  def clear_socket_buffer(gripper_socket="1", read_timeout = 0.1):
      rq_comm_clear_socket_buffer_enabled[rq_socket_to_index(gripper_socket)] = True
  end

  def rq_gripper_id_to_ascii(gripper_id):
      if(gripper_id == "1"):
          return 57
      elif(gripper_id == "2"):
          return 50
      elif(gripper_id == "3"):
          return 51
      elif(gripper_id == "4"):
          return 52
      end
  end

      def scale(value, rawRange, scaledRange):
          def computeSlope(inputRange, outputRange):
              outputRangeDelta = outputRange[1] - outputRange[0]
              inputRangeDelta = inputRange[1] - inputRange[0]

              if (inputRangeDelta == 0):
                  return 0
              else:
                  return outputRangeDelta / inputRangeDelta
              end
          end

          def computeIntercept(slope, inputRange, outputRange):
              return outputRange[0] - (slope * inputRange[0])
          end

          def clipScaledValue(outputScaledValue, outputRange):
              if (outputRange[0] < outputRange[1]):
                  return clipWhenLowerLimitIsLessThanHigher(outputScaledValue, outputRange)
              else:
                  return clipWhenLowerLimitIsGreaterThanHigherLimit(outputScaledValue, outputRange)
              end
          end

          def clipWhenLowerLimitIsGreaterThanHigherLimit(outputScaledValue, outputRange):
              if (outputScaledValue < outputRange[1]):
                  return outputRange[1]
              elif (outputScaledValue > outputRange[0]):
                  return outputRange[0]
              else:
                  return outputScaledValue
              end
          end

          def clipWhenLowerLimitIsLessThanHigher(outputScaledValue, outputRange):
              if (outputScaledValue < outputRange[0]):
                  return outputRange[0]
              elif (outputScaledValue > outputRange[1]):
                  return outputRange[1]
              else:
                  return outputScaledValue
              end
          end

          slope = computeSlope(rawRange, scaledRange)
          intercept = computeIntercept(slope, rawRange, scaledRange)
          scaledValue = slope * value + intercept
          return clipScaledValue(scaledValue, scaledRange)
      end

      def limit(value, range):
          return scale(value, range, range)
      end


  rq_init_comm_if_connected(9, "1")
  rq_init_comm_if_connected(2, "2")
  rq_init_comm_if_connected(3, "3")
  rq_init_comm_if_connected(4, "4")
  rq_print_connected_grippers()
  rq_gripper_communication_thread = run rq_gripper_communication()
  set_closed_norm(97.6470588235294, "1")
  set_open_norm(1.1764705882352942, "1")
  set_closed_mm(0.0, "1")
  set_open_mm(53.0, "1")
  set_closed_norm(100.0, "2")
  set_open_norm(0.0, "2")
  set_closed_mm(0.0, "2")
  set_open_mm(50.0, "2")
  set_closed_norm(100.0, "3")
  set_open_norm(0.0, "3")
  set_closed_mm(0.0, "3")
  set_open_mm(50.0, "3")
  set_closed_norm(100.0, "4")
  set_open_norm(0.0, "4")
  set_closed_mm(0.0, "4")
  set_open_mm(50.0, "4")
  rq_current_limit_enabled = False
  while(not rq_gripper_communication_thread_started):
      sleep(0.008)
  end
  # end: URCap Installation Node
  global AMR_Position=struct(position_identifier=0, x1=0, x2=0, y1=0, y2=0, theta1=0, theta2=0)
  global CAM_Pose=p[0,0,0,0,0,0]
  global CAM_Relation=""
  global CMD_Abort=  False
  global CMD_Clear=  False
  global CMD_Reset=  False
  global CMD_Start=  False
  global CMD_Suspend=  False
  global CMD_Unhold=  False
  global CMD_Unsuspend=  False
  global CNT_Rack_Output=0
  global FNC_Freedrive=  False
  global PRC_TubCounter=0
  global STP=0
  global easyPickCount_4=0
  global easyPickCount_7=0
  global easyPickNoObj_4=0
  global easyPickNoObj_7=0
  global easyPickParts_4=0
  global easyPickParts_7=0
  global TMR_Barcode=0
  global Container_mid_1_p=p[-.379239199143, -.127191311915, .299999999998, .000000000046, -.000000000021, -1.247199999994]
  global Container_mid_1_q=[-2.477408934449926, -1.2969853503591224, -1.875639182904262, -1.539621866126728, 1.5731943360401213, -2.8009955944022717]
  global trigger_otw_p=p[-.364831738276, -.163967193938, .343299997821, .000000000046, -.000000000020, -1.148401333327]
  global trigger_otw_q=[-2.378283213085033, -1.2994862387706814, -1.7634300687554951, -1.6493302004167063, 1.573123683454141, -2.8011223671816943]
  global Waypoint_54_p=p[.008800512419, -.547926542621, .402696567415, -.589884378425, -.007228654778, -.061268144704]
  global Waypoint_54_q=[-1.2044575850116175, -1.3416667741588135, -1.8272563219070435, -0.9884541195682068, 1.3621035814285278, -2.7712565104113978]
  global Waypoint_77_p=p[-.178371829612, -.433927395311, .368082383916, -.086593488055, .704679941724, -.007869906074]
  global Waypoint_77_q=[-1.265390698109762, -1.3355963987163086, -1.7944865226745605, -1.7402602634825648, 0.8780410885810852, -2.7713127771960657]
  global Waypoint_83_p=p[.008800512419, -.547926542621, .402696567415, -.589884378425, -.007228654778, -.061268144704]
  global Waypoint_83_q=[-1.2044575850116175, -1.3416667741588135, -1.8272563219070435, -0.9884541195682068, 1.3621035814285278, -2.7712565104113978]
  global Waypoint_84_p=p[-.178371829612, -.433927395311, .368082383916, -.086593488055, .704679941724, -.007869906074]
  global Waypoint_84_q=[-1.265390698109762, -1.3355963987163086, -1.7944865226745605, -1.7402602634825648, 0.8780410885810852, -2.7713127771960657]
  global Vial_above_1_p=p[.017105793010, -.652093028359, .184920586844, .000000000272, .000000000270, 1.564063451276]
  global Vial_above_1_q=[-1.3375440709712851, -1.9618096977868804, -1.4665759083780685, -1.2837941559171444, 1.5732503672317195, -4.47276330421513]
  global Vial_pick_poi_1_p=p[.017105792852, -.648922724010, .093307568731, .000000000271, .000000000270, 1.564063451276]
  global Vial_pick_poi_1_q=[-1.3366329456391917, -2.0375277831965413, -1.6071432798879028, -1.0675084332049813, 1.57309887265915, -4.471135348858068]
  global Waypoint_86_p=p[.019227646885, -.648669633640, .184920586950, .000000000000, .000000000000, .024063451426]
  global Waypoint_86_q=[-1.3331129109407733, -1.9540750545686123, -1.4775914902901128, -1.280581784992414, 1.5733500744865856, -2.928303704452631]
  global Waypoint_87_p=p[-.032361834699, -.348336136197, .391475576335, -.000008499254, .000014589902, -.004651426820]
  global Waypoint_87_q=[-1.2709335019096129, -1.1914598663441005, -1.708995335060501, -1.8117888533498316, 1.5729683532263925, -2.8379347397710237]
  global Vial_3FG_plac_1_p=p[-.031858676359, -.349402499566, .145301120695, .000000000000, .000000000000, .000000000000]
  global Vial_3FG_plac_1_q=[-1.2723975525801707, -1.252376585823825, -2.3128114007049496, -1.1470592278900167, 1.5730548099411423, -2.8414815174610535]
  global Waypoint_88_p=p[-.032361834699, -.348336136197, .391475576335, -.000008499254, .000014589902, -.004651426820]
  global Waypoint_88_q=[-1.2709335019096129, -1.1914598663441005, -1.708995335060501, -1.8117888533498316, 1.5729683532263925, -2.8379347397710237]
  global cap_dump_1_p=p[-.139168676487, -.420163541420, .146096395183, .000000000000, .000000000000, .000000000000]
  global cap_dump_1_q=[-1.584588644510994, -1.5093464179777323, -2.1118449369620347, -1.091059703602438, 1.5728943834877336, -3.154014906686923]
  global Waypoint_89_p=p[-.032361834699, -.348336136197, .391475576335, -.000008499254, .000014589902, -.004651426820]
  global Waypoint_89_q=[-1.2709335019096129, -1.1914598663441005, -1.708995335060501, -1.8117888533498316, 1.5729683532263925, -2.8379347397710237]
  global Vial_3FG_plac_2_p=p[-.031858676359, -.349402499566, .145301120695, .000000000000, .000000000000, .000000000000]
  global Vial_3FG_plac_2_q=[-1.2723975525801707, -1.252376585823825, -2.3128114007049496, -1.1470592278900167, 1.5730548099411423, -2.8414815174610535]
  global Waypoint_90_p=p[-.032361834699, -.348336136197, .391475576335, -.000008499254, .000014589902, -.004651426820]
  global Waypoint_90_q=[-1.2709335019096129, -1.1914598663441005, -1.708995335060501, -1.8117888533498316, 1.5729683532263925, -2.8379347397710237]
  global cap_dump_2_p=p[-.139168676487, -.420163541420, .146096395183, .000000000000, .000000000000, .000000000000]
  global cap_dump_2_q=[-1.584588644510994, -1.5093464179777323, -2.1118449369620347, -1.091059703602438, 1.5728943834877336, -3.154014906686923]
  global Waypoint_91_p=p[-.032361834699, -.348336136197, .391475576335, -.000008499254, .000014589902, -.004651426820]
  global Waypoint_91_q=[-1.2709335019096129, -1.1914598663441005, -1.708995335060501, -1.8117888533498316, 1.5729683532263925, -2.8379347397710237]
  global Vial_liq_abov_1_p=p[-.025303660977, -.338758622354, .426628485936, -1.315858642253, .800043520260, -.928295855026]
  global Vial_liq_abov_1_q=[-0.3789628187762659, -1.5149522957256814, -2.263045310974121, 0.7870649534412841, -0.750984017048971, -3.2237566153155726]
  global Vial_liq_pick_3_p=p[-.002660428945, -.335984893034, .159389832934, -1.150456778400, .673175527684, -1.010612657503]
  global Vial_liq_pick_3_q=[-0.3660772482501429, -1.4503649038127442, -2.4056053161621094, -1.994692941705221, 0.8039668202400208, -0.2508929411517542]
  global Vial_liq_pick_4_p=p[-.041402486291, -.356791603314, .125395323246, -1.143483969075, .651070210027, -.878721885453]
  global Vial_liq_pick_4_q=[-0.4426233705502476, -1.437252121513727, -2.551930962114307, -1.776528229806984, 0.6562026234073748, -0.43018811960029524]
  global Vial_liq_abov_2_p=p[-.025303660977, -.338758622354, .426628485936, -1.315858642253, .800043520260, -.928295855026]
  global Vial_liq_abov_2_q=[-0.3789628187762659, -1.5149522957256814, -2.263045310974121, 0.7870649534412841, -0.750984017048971, -3.2237566153155726]
  global Liquid_midway_1_p=p[.057575295009, -.583081747994, .306414980749, -1.351675548728, .120935756539, -.096908606303]
  global Liquid_midway_1_q=[-0.895174805318014, -1.7035466633238734, -2.380953073501587, 0.631549521083496, 0.7706599235534668, -2.9455552736865442]
  global shake_3_p=p[.057574880217, -.583085370269, .306422893466, -1.360996190983, -.155555042453, -.438136255921]
  global shake_3_q=[-0.8951800505267542, -1.7035466633238734, -2.380937099456787, 0.6315542894550782, 0.7706599235534669, -2.5394540616517496]
  global shake_4_p=p[.057581636113, -.583090570002, .306439684073, -1.308767904323, .368530312677, .214926493520]
  global shake_4_q=[-0.8951714674579065, -1.7035395107665003, -2.380906343460083, 0.6315504747578125, 0.7706480026245118, -3.3161255787892268]
  global drop_above_3_p=p[.268235025993, -.467784390499, .226219872376, -1.027832627524, -.430841408251, 1.004603115937]
  global drop_above_3_q=[-0.935645882283346, -1.6663371525206507, -2.4252893924713135, 0.41966931402172847, 1.8470635414123535, -3.4600217978106897]
  global drop_above_4_p=p[.219042229014, -.470775657081, .133754190740, -.313004595901, -.344395319364, 1.500564994056]
  global drop_above_4_q=[-1.0601594887284795, -1.70046459045642, -2.0799996233759863, -0.7243227230676759, 1.9429634314685202, -4.115129153870795]
  global liq_tran_3_p=p[.213067510942, -.469567035397, .100231043184, .251862243732, .217902579404, 1.592812335393]
  global liq_tran_3_q=[-0.7789645168037476, -1.822364827406652, -1.8643518410805573, -1.252158963840138, 1.3768134449520435, -3.9328333233290254]
  global drop_above_5_p=p[.219042229014, -.470775657081, .133754190740, -.313004595901, -.344395319364, 1.500564994056]
  global drop_above_5_q=[-1.0601594887284795, -1.70046459045642, -2.0799996233759863, -0.7243227230676759, 1.9429634314685202, -4.115129153870795]
  global Waypoint_92_p=p[.187119460405, -.493959476151, .133754190608, -.313004596540, -.344395317757, 1.500564993991]
  global Waypoint_92_q=[-1.1418328121400876, -1.7310553375189475, -2.033634768766424, -0.772026910513711, 1.958578934631971, -4.201588449364511]
  global liq_tran_4_p=p[.195957706507, -.493022614126, .100231042689, .160718757180, .109807038912, 1.525321508623]
  global liq_tran_4_q=[-0.881740380645474, -1.8244526267589851, -1.865100964490387, -1.1608866323693583, 1.4631433601076713, -3.973915130363038]
  global drop_above_6_p=p[.219042229014, -.470775657081, .133754190740, -.313004595901, -.344395319364, 1.500564994056]
  global drop_above_6_q=[-1.0601594887284795, -1.70046459045642, -2.0799996233759863, -0.7243227230676759, 1.9429634314685202, -4.115129153870795]
  global drop_above_7_p=p[.268235025993, -.467784390499, .226219872376, -1.027832627524, -.430841408251, 1.004603115937]
  global drop_above_7_q=[-0.935645882283346, -1.6663371525206507, -2.4252893924713135, 0.41966931402172847, 1.8470635414123535, -3.4600217978106897]
  global Liquid_midway_2_p=p[.057575295009, -.583081747994, .306414980749, -1.351675548728, .120935756539, -.096908606303]
  global Liquid_midway_2_q=[-0.895174805318014, -1.7035466633238734, -2.380953073501587, 0.631549521083496, 0.7706599235534668, -2.9455552736865442]
  global Vial_drop_abo_1_p=p[.000324902251, -.648569523142, .221894115667, -.873462921366, 1.165852672573, -1.482720593185]
  global Vial_drop_abo_1_q=[-1.0576906334721352, -2.393016994184633, -0.9236232851859159, -2.5729213042279273, 0.7903331288549689, -0.33286325848155585]
  global Vial_liq_drop_1_p=p[.001020867953, -.647659915585, .092915870838, -.834762611599, 1.081942994823, -1.540647900176]
  global Vial_liq_drop_1_q=[-1.0631954168193474, -2.4447642951220825, -1.128811017825127, -2.1983115491972294, 0.8130148661460634, -0.38984988696911316]
  global Vial_drop_abo_2_p=p[.000324902251, -.648569523142, .221894115667, -.873462921366, 1.165852672573, -1.482720593185]
  global Vial_drop_abo_2_q=[-1.0576906334721352, -2.393016994184633, -0.9236232851859159, -2.5729213042279273, 0.7903331288549689, -0.33286325848155585]
  global Spatula_otw_p=p[-.038472058237, -.263141484147, .425351216717, -.000441582511, -.000128175490, 3.034387645854]
  global Spatula_otw_q=[-1.1888947506684495, -1.0083288774886814, -1.7052227056065874, -1.9984805067363443, 1.5730180972985317, 0.48793409320312264]
  global pick_spat_L_abv_p=p[.239059466375, -.067212518441, .280720723617, .000017217488, -.000484427718, 3.106837214660]
  global pick_spat_L_abv_q=[0.292765616142962, -0.8565557553273315, -2.140199892763044, -1.715349495646084, 1.573623142106424, 1.8984976776985687]
  global spat_L_pick_p=p[.242468789885, -.067301915011, .193171208067, .000017217488, -.000484427718, 3.106837214657]
  global spat_L_pick_q=[0.2867414378807389, -0.8600077002089179, -2.3629148016312627, -1.4891831672860159, 1.5737695566221115, 1.8933890858591198]
  global spat_L_lift_p=p[.245402002494, -.067432373551, .289049296496, .000017217490, -.000484427724, 3.106837214657]
  global spat_L_lift_q=[0.2834351187564135, -0.8798320076811592, -2.1119436738532986, -1.7203314352121302, 1.573588313403067, 1.8891054681654005]
  global spat_L_side_p=p[.247133573905, -.017633681797, .289062935631, .000017217490, -.000484427724, 3.106837214657]
  global spat_L_side_q=[0.49719173575848863, -0.8582398211168538, -2.1182130454788215, -1.735610316654931, 1.5735817737572706, 2.1028402698705397]
  global spat_L_up_p=p[.247135508752, -.017665230822, .397130746165, .000017217490, -.000484427724, 3.106837214657]
  global spat_L_up_q=[0.49854946074076967, -0.9346239623559676, -1.808280269374471, -1.969158816463132, 1.5731020084036995, 2.1031742024348157]
  global spat_M_up_p=p[.244670000000, -.112000000000, .420343789747, .000026293990, -.000477463070, 3.067686800857]
  global spat_M_up_q=[0.09097498152209688, -1.0114245603211778, -1.718034632879454, -1.9826932847219538, 1.5730130135866505, 1.734554438783734]
  global spat_M_pick_p=p[.244673518506, -.111985070134, .192299022723, .000043885692, -.000001622442, 3.067686841404]
  global spat_M_pick_q=[0.08868170265231701, -0.9271392933223233, -2.343826449241451, -1.441236864368305, 1.5733923850045939, 1.7345552462242537]
  global spat_S_Up_7_p=p[.243228810603, -.161948321982, .423281604617, .000026293955, -.000477463064, 3.067686800854]
  global spat_S_Up_7_q=[-0.11182322368059516, -1.0716267311491734, -1.6854498186860427, -1.955120134033855, 1.5730106579635699, 1.5317349120701778]
  global spat_S_Pick_4_p=p[.245377020686, -.158668022535, .192285730279, .000026293985, -.000477463062, 3.067686800840]
  global spat_S_Pick_4_q=[-0.10087203759495189, -1.011188488703386, -2.311978084495874, -1.3890267520590838, 1.5735990551056096, 1.5450562970948172]
  global spat_S_Up_8_p=p[.252087445596, -.159242094834, .423281604617, .000026293954, -.000477463070, 3.067686800855]
  global spat_S_Up_8_q=[-0.09804692328730358, -1.0862987822056382, -1.6788706463996483, -1.9470242450550348, 1.5730147401359813, 1.5455107082823842]
  global spat_flatM_up_p=p[.229022666361, -.211442909333, .418634047126, .000026293953, -.000477463083, 3.067686800888]
  global spat_flatM_up_q=[-0.30183372580416545, -1.1157042924275036, -1.6775646144685776, -1.9189678841796578, 1.5730340557943228, 1.341766142011193]
  global spat_flatM_pick_p=p[.241028983327, -.208057297586, .192270533170, .000026293950, -.000477463079, 3.067686800885]
  global spat_flatM_pick_q=[-0.2805687960562633, -1.1003763929487214, -2.271431297337675, -1.3404236887924883, 1.5734924238720627, 1.3653813047742556]
  global spat_flatS_up_p=p[.237651953780, -.253943828614, .403961222825, .000026293950, -.000477463092, 3.067686800841]
  global spat_flatS_up_q=[-0.42363550926974103, -1.1939944599502539, -1.6745915127240307, -1.843675057902054, 1.5731001874678698, 1.220082820532415]
  global spat_flatS_pick_p=p[.241325662334, -.251726327528, .192256842740, .000026293947, -.000477463087, 3.067686800841]
  global spat_flatS_pick_q=[-0.4144907797170738, -1.1967447109013012, -2.21926362252748, -1.2962499335425761, 1.5733885098427622, 1.2314402238866728]
  global spat_S_pick_p=p[.238158866340, -.157926795425, .192632100345, .000026293989, -.000477463069, 3.067686800857]
  global spat_S_pick_q=[-0.10084756991493293, -0.9881392730064915, -2.3204232610157494, -1.403630829593915, 1.5736254260650586, 1.5450653591083503]
  global spat_S_up_p=p[.244260523725, -.164466690315, .417087579736, .000026293988, -.000477463072, 3.067686800857]
  global spat_S_up_q=[-0.12101499604198729, -1.0718307017854336, -1.7023391702814736, -1.938028805938881, 1.573044424728474, 1.5226045951991447]
  global Waypoint_7_p=p[-.472820924474, .292439826233, .207418370237, -.137787250486, 2.177332259632, -2.152029714756]
  global Waypoint_7_q=[-2.911134078210732, -1.90240864358569, -1.968768330510411, -2.500365101593811, 0.11427687110891149, 0.0958980389250167]
  global Waypoint_8_p=p[-.357612884176, -.251084817998, .212379799667, -.858181193174, 1.714832512191, -1.687547565568]
  global Waypoint_8_q=[-1.620834863369681, -1.8936194567376496, -1.9821394403832038, -2.4599791457905273, 0.6296693672615152, 0.07625365420707819]
  global Decapp_above_3_p=p[-.013480295948, -.359153355979, .266194408367, -.879653555922, 1.646336924805, -1.709111068605]
  global Decapp_above_3_q=[-0.9632157249872035, -2.0163405763031657, -1.5968194594157152, -2.6579215719847085, 1.251243398585566, 0.047906446502667066]
  global Decapp_place_3_p=p[-.013480295890, -.359153356055, .160907502384, -.879653554902, 1.646336919740, -1.709111066456]
  global Decapp_place_3_q=[-0.9633402410919709, -2.1541179572356635, -1.6937729380888573, -2.4232786481058053, 1.2517342187662468, 0.04818402956922263]
  global Decapp_above_4_p=p[-.013480295948, -.359153355979, .266194408367, -.879653555922, 1.646336924805, -1.709111068605]
  global Decapp_above_4_q=[-0.9632157249872035, -2.0163405763031657, -1.5968194594157152, -2.6579215719847085, 1.251243398585566, 0.047906446502667066]
  global Waypoint_78_p=p[-.051450028091, -.519555688329, .365718563414, -1.287302938145, 1.077637394477, -1.218524965834]
  global Waypoint_78_q=[-0.9214276262416012, -1.8899696965062578, -1.4939326452510562, -2.840015661555725, 0.5585157189668353, 0.033997638875617575]
  global Waypoint_10_p=p[-.330595116596, .282932669854, .220236276291, 1.304675539882, .014233792938, -1.753932442581]
  global Waypoint_10_q=[-3.189526379253601, -1.8418198435143305, -1.7138504750370807, -2.182789974066381, 1.0126080912871243, -2.4455984844694645]
  global Waypoint_9_p=p[-.538777454962, .370695704977, .175030018143, -.317104215445, 2.082346543003, -2.037631421082]
  global Waypoint_9_q=[-3.1158871966457857, -1.998548595120492, -1.941797010061462, -2.2703530575838844, -0.27573365931009164, -0.06926782177267654]
  global Powder_wayp1_p=p[-.472820924474, .292439826233, .207418370237, -.137787250486, 2.177332259632, -2.152029714756]
  global Powder_wayp1_q=[-2.911134078210732, -1.90240864358569, -1.968768330510411, -2.500365101593811, 0.11427687110891149, 0.0958980389250167]
  global Waypoint_2_p=p[-.357612884176, -.251084817998, .212379799667, -.858181193174, 1.714832512191, -1.687547565568]
  global Waypoint_2_q=[-1.620834863369681, -1.8936194567376496, -1.9821394403832038, -2.4599791457905273, 0.6296693672615152, 0.07625365420707819]
  global Postions_otw_p=p[-.010896578244, -.533368729951, .288851175116, -1.233738470894, 1.195331112012, -1.207314088469]
  global Postions_otw_q=[-0.898791023514228, -2.078490033037677, -1.4499891355755317, -2.7624416226992476, 0.6570218891920963, 0.02136606178275929]
  global cont_A_otw_p=p[.070238108556, -.655257851554, .184611566008, -1.090601381517, 1.404822685081, -1.413645380264]
  global cont_A_otw_q=[-0.990969136335913, -2.7123780097559784, -0.5772671651193146, -3.0005537851220403, 0.84719335943793, 0.020652463706785973]
  global cont_B_otw_p=p[.255895686750, -.501120003087, .157855243207, -1.209177187561, 1.209243088037, -1.209202949417]
  global cont_B_otw_q=[-0.5819602570351563, -2.5181180937953833, -1.0264696604583161, -2.7360726814058687, 0.9880932038785559, -0.004134033524621827]
  global cont_B_safe_p=p[.242897168204, -.501733713795, .237745474779, -1.209212324107, 1.209144328638, -1.209309913894]
  global cont_B_safe_q=[-0.5929699566143585, -2.4210115429142114, -0.9949203644592259, -2.8646436479104267, 0.976678899749076, -0.004020526358775811]
  global cont_C_otw_p=p[.319495487998, -.362719410364, .163846736977, -1.233784872294, 1.195277203291, -1.207325031551]
  global cont_C_otw_q=[-0.3611889651645974, -2.404603865546651, -1.2341573845076566, -2.650535279811077, 1.1944844573128257, 0.01638086594640864]
  global Waypoint_1_p=p[-.352029261722, -.424157832422, .472326578019, -.000004407962, .000020663369, -1.529709227737]
  global Waypoint_1_q=[-2.017015745614491, -1.7423968528991196, -1.0053357238485425, -1.9644715035904907, 1.5727249689896, -2.060727852912713]
  global Waypoint_5_p=p[.219993437017, -.447144142811, .462350040687, .000006087494, .000031090075, .000022232405]
  global Waypoint_5_q=[-0.8406239476037944, -1.5982534362206806, -1.1934200873248484, -1.9205794898315975, 1.5727336676986443, -2.4135960466995314]
  global place_2_home_p=p[-.352029261717, -.424157832411, .329197314759, -.000004407962, .000020663369, -1.529709227737]
  global place_2_home_q=[-2.017880982348384, -1.6708952803108668, -1.462293789471877, -1.5790150659586653, 1.5732060241635952, -2.059940179665328]
  global PosA_up_p=p[.028578953747, -.638006009765, .227275735849, -1.090660933958, 1.404791542934, -1.413645191233]
  global PosA_up_q=[-1.0254743496427432, -2.565176838504783, -0.7558042274983681, -2.9696064674274343, 0.8129191411995651, 0.021444818458024387]
  global PosA_pick_p=p[.026918718687, -.640084889741, .097901147521, -1.090660933959, 1.404791542934, -1.413645191233]
  global PosA_pick_q=[-1.028821435558534, -2.6899890636403807, -0.8526126047665157, -2.7478942693937167, 0.8103607002888742, 0.021326778146411485]
  global PosB_up_p=p[.239472634782, -.492481416782, .220767759213, -1.233738470883, 1.195331111998, -1.207314088469]
  global PosB_up_q=[-0.5800230603397054, -2.4076296700885997, -1.0699783327330836, -2.8116344407747427, 0.9750472858169287, 0.017627507888886562]
  global PosB_pick_p=p[.240630296955, -.494558620171, .096392895280, -1.233740573549, 1.195309876041, -1.207293779132]
  global PosB_pick_q=[-0.5816146260408139, -2.553273721769836, -1.1376320925804277, -2.5983292591462153, 0.9740936784345416, 0.017625262979849232]
  global PosC_up_p=p[.241566602786, -.359249123455, .230260583862, -1.233738470888, 1.195331111997, -1.207314088449]
  global PosC_up_q=[-0.39573787962534546, -2.2019009616581497, -1.4115270142506517, -2.675987785326166, 1.160180741930842, 0.01687917643039505]
  global PosC_pick_p=p[.240633854030, -.361553124916, .093979792658, -1.233738470878, 1.195331111997, -1.207314088469]
  global PosC_pick_q=[-0.39992427526118757, -2.386042391328985, -1.4894374567278712, -2.414022930893381, 1.1566786195951169, 0.01712017454263659]
  global Pow_decap_up_p=p[-.017556487132, -.367519866742, .275835445416, -.605635182849, 1.892518157522, -1.890848751165]
  global Pow_decap_up_q=[-1.1272088681128203, -2.1173924123331025, -1.4250048354055203, -2.7485980486387676, 1.4193896902217862, 0.023247957637719453]
  global pow_decap_place_p=p[-.020433194420, -.368310202914, .161281291611, -.605635182838, 1.892518157522, -1.890848751163]
  global pow_decap_place_q=[-1.132360890531647, -2.2521863255983092, -1.5302136899970318, -2.5086176644751683, 1.4149282844269635, 0.02347140074572661]
  global Decap_above_p=p[-.031863883354, -.349974838955, .288042264213, .000000000000, .000000000000, .000000000000]
  global Decap_above_q=[-1.271900116540503, -1.1670201114602632, -1.989291655468758, -1.5559360538518163, 1.573255119759632, -2.842476569674073]
  global Decapp_p=p[-.031864263150, -.349974612700, .230259377740, .000000000000, .000000000000, .000000000000]
  global Decapp_q=[-1.2723555431601419, -1.1810456878410935, -2.1291754890757737, -1.4020263844320349, 1.5732701843074919, -2.842325632263757]
  global Cap_above_p=p[-.224192409203, -.629599568633, .257274081142, .000015605575, -.000015166009, -1.647823825902]
  global Cap_above_q=[-1.710642681834492, -1.9674285251810462, -1.2705185053146897, -1.4742193161331247, 1.573506065067499, -1.6347709465008595]
  global Cap_place_p=p[-.224189049846, -.629597879697, .041885651757, .000015605572, -.000015166011, -1.647823825903]
  global Cap_place_q=[-1.7111696563854295, -2.13979870939016, -1.5941008764912503, -0.978265561728648, 1.5732789016410962, -1.6336328794662904]
  global OP_PowderA2_p=p[.009371277507, -.409434369247, .294169017766, -.823281033205, 1.709410851243, -1.698303593897]
  global OP_PowderA2_q=[-0.9994544761745754, -2.1395254572673217, -1.3437567783153916, -2.8143375616690456, 1.2617899549595724, 0.019614613715634555]
  global Decap_up_p=p[-.018339217391, -.367674469480, .249553854268, -.546164737599, 1.935964719000, -1.930057109666]
  global Decap_up_q=[-1.158124747223252, -2.1569920012936787, -1.4340832185069745, -2.7006032680036753, 1.4556626828962336, 0.02060977878679182]
  global Decap_pick_p=p[-.020429098827, -.367971872627, .161604333799, -.546164737600, 1.935964719000, -1.930057109666]
  global Decap_pick_q=[-1.161653098289774, -2.263509236689538, -1.5087211318402236, -2.519459740767391, 1.452646640403743, 0.02077912034002202]
  global Op_PowA_wP_p=p[-.173727579245, -.372934016396, .295116627479, -.972390492433, 1.540962074418, -1.548745344994]
  global Op_PowA_wP_q=[-1.1740587397768483, -1.865656321049359, -1.7426943793777419, -2.679427276872525, 0.8588908769087338, 0.017944699631825187]
  global Waypoint_12_p=p[-.812560029877, -.415067232840, .258518340146, -1.257569567036, 1.159670338548, -1.145019586130]
  global Waypoint_12_q=[-2.3224548809497123, -2.3211405271930765, -1.1304722687551445, -2.8155296475017018, -0.8321758827962036, -0.007205995478960503]
  global Waypoint_18_p=p[-.813643087636, -.416224939441, .090971414301, -1.257570310932, 1.159676546329, -1.145010619026]
  global Waypoint_18_q=[-2.3224916967547475, -2.513993544062452, -1.2408975037093848, -2.5121717481246186, -0.831286599209303, -0.007326414722441221]
  global Waypoint_19_p=p[-.812560029269, -.415067232191, .079455005744, -1.257569567033, 1.159670338546, -1.145019586137]
  global Waypoint_19_q=[-2.3224951834453367, -2.5274729453886575, -1.2489176533831348, -2.4906644180980346, -0.8312252662037514, -0.007338111970053518]
  global TMR_Barcode_is_counting=False
  thread Timer_Thread():
    while (True):
      if (TMR_Barcode_is_counting):
        TMR_Barcode = TMR_Barcode + get_steptime()
      end
      sync()
    end
  end
  run Timer_Thread()
  def Sub_Vision_V18():
    $ 847 "Sub_Vision_V18" "noBreak"
    $ 848 "PreSettings"
    $ 849 "CAM_LM_Detected≔ False "
    global CAM_LM_Detected=  False
    $ 850 "CAM_Captures≔0"
    global CAM_Captures=0
    $ 851 "CAM_Pose≔p[0,0,0,0,0,0]"
    global CAM_Pose=p[0,0,0,0,0,0]
    $ 852 "CAM_LM_Refinmnt≔ False "
    global CAM_LM_Refinmnt=  False
    $ 853 "CAM_LM_Refined≔ False "
    global CAM_LM_Refined=  False
    $ 854 "CAM_LM_Deviatn≔p[0,0,0,0,0,0]"
    global CAM_LM_Deviatn=p[0,0,0,0,0,0]
    $ 855 "CAM_LM_ID≔0"
    global CAM_LM_ID=0
    $ 856 "CAM_Done≔ False "
    global CAM_Done=  False
    $ 857 "CAM_CNT_Obj≔0"
    global CAM_CNT_Obj=0
    $ 858 "CAM_Result = []"
    CAM_Result = []
    $ 859 "OBJ_Detected≔ False "
    global OBJ_Detected=  False
    $ 860 "FRM_Reference≔p[0,0,0,0,0,0]"
    global FRM_Reference=p[0,0,0,0,0,0]
    $ 861 "'=========='"
    # '=========='
    $ 862 "Switch Action"
    switch_1 = Action
    $ 863 "Case 13"
    if (13 == switch_1):
    elif (15 == switch_1):
      $ 981 "Case 15"
    elif (131 == switch_1):
      $ 1027 "Case 131"
      $ 1028 "Read (SensoPart)"
      $ 1029 "Action_Info≔'search for landmark'"
      global Action_Info="search for landmark"
      $ 1030 "CAM_LM≔CAM_LMs[4]"
      global CAM_LM=CAM_LMs[4]
      $ 1031 "CAM_Relation≔CAM_LM.capture_relation"
      global CAM_Relation=CAM_LM.capture_relation
      $ 1032 "go to capture pose"
      $ 1035 "If ITM_ID≟1 and JIG≟7"
      if (ITM_ID == 1  and  JIG == 7):
        $ 1036 "PSE_T≔uLM_Cap_SSRack"
        global PSE_T=uLM_Cap_SSRack
      else:
        $ 1037 "ElseIf ITM_ID≟5 and JIG≟7"
        if (ITM_ID == 5  and  JIG == 7):
          $ 1038 "PSE_T≔FRM_Cap_SSRack"
          global PSE_T=FRM_Cap_SSRack
        else:
          $ 1041 "ElseIf ITM_ID≟1 and JIG≟15"
          if (ITM_ID == 1 and JIG == 15):
            $ 1042 "MoveJ"
            $ 1043 "Container_mid_1" "breakAfter"
            movej(get_inverse_kin(Container_mid_1_p, qnear=Container_mid_1_q), a=1.3962634015954636, v=1.0471975511965976, r=0.05)
            $ 1045 "PSE_T≔FRM_Container_const"
            global PSE_T=p[-0.5003348223692186,0.35061804815168285,0.41579001388808423,-5.092943187272062E-5,1.0145185065363121E-4,-2.764319258713288]
          else:
            $ 1046 "ElseIf ITM_ID≟1 and JIG≟21"
            if (ITM_ID == 1 and JIG == 21):
              $ 1048 "PSE_T≔FRM_PoTS_const"
              global PSE_T=p[-0.5403054403210852,-0.10910773999775857,0.4828,3.058497512721046E-6,2.3454853329357316E-5,-2.208510541952706]
            else:
              $ 1049 "ElseIf ITM_ID≟1 and JIG≟17"
              if (ITM_ID == 1 and JIG == 17):
                $ 1050 "MoveJ"
                $ 1051 "zero_scale()"
                zero_scale()
                $ 1052 "trigger_otw" "breakAfter"
                movej(get_inverse_kin(trigger_otw_p, qnear=trigger_otw_q), a=1.3962634015954636, v=1.0471975511965976, r=0.05)
                $ 1056 "PSE_T≔FRM_weigh_scale_const"
                global PSE_T=p[-0.3804866881697204,0.025744252835212,0.4723487455232425,-1.0445769542396123E-4,-1.924788411074358E-5,-2.1691978730572363]
              end
            end
          end
        end
      end
      $ 1057 "do_transition(PSE_T, keep_rxry=False)"
      do_transition(PSE_T, keep_rxry=False)
      $ 1058 "Set"
      set_tcp(p[0.0,0.0,0.161,3.1415,0.0,0.0])
      $ 1059 "MoveJ"
      $ 1060 "PSE_T" "breakAfter"
      movej(PSE_T, a=1.3962634015954636, v=1.7453292519943295)
      $ 1061 "CAM_Pose≔get_actual_tcp_pose()"
      global CAM_Pose= get_actual_tcp_pose ()
      $ 1062 "Loop  not CAM_Done and  not ERROR.FLAG and  not CMD_Stop"
      while (  not  CAM_Done  and    not  ERROR.FLAG  and    not  CMD_Stop):
        $ 1063 "adjust capture pose"
        $ 1064 "If CAM_LM_Detected and CAM_LM_Refinmnt"
        if (CAM_LM_Detected  and  CAM_LM_Refinmnt):
          $ 1065 "PSE_T≔p[0,0,0.300,0,0,0]"
          global PSE_T=p[0,0,0.300,0,0,0]
          $ 1066 "CAM_Pose≔PSE_T"
          global CAM_Pose=PSE_T
          $ 1067 "If  not is_reachable(FRM_Reference,[PSE_T])"
          if (  not  is_reachable(FRM_Reference,[PSE_T])):
            $ 1068 "Error"
            $ 1069 "set_error(ERROR_POSE_NOT_REACHABLE)"
            set_error(ERROR_POSE_NOT_REACHABLE)
          end
          $ 1070 "If  not ERROR.FLAG"
          if (  not  ERROR.FLAG):
            $ 1071 "MoveJ"
            $ 1072 "PSE_T" "breakAfter"
            set_tcp(p[0.0,0.0,0.161,0.0,0.0,0.0])
            movej(pose_trans(FRM_Reference, PSE_T), a=0.8726646259971648, v=1.3962634015954636)
            $ 1073 "CAM_LM_Refined≔ True "
            global CAM_LM_Refined=  True
          end
        else:
          $ 1074 "ElseIf  not CAM_LM_Detected and CAM_Captures>0"
          if (  not  CAM_LM_Detected  and  CAM_Captures>0):
            $ 1075 "MoveL"
            $ 1076 "If FRM_Reference≟p[0,0,0,0,0,0]"
            if (FRM_Reference == p[0,0,0,0,0,0]):
              $ 1077 "PSE_T≔get_random_pose(pose_ref=CAM_Pose, mode='cubic', range_max=[0.150,0.150,0.015])"
              global PSE_T=get_random_pose(pose_ref=CAM_Pose, mode="cubic", range_max=[0.150,0.150,0.015])
            else:
              $ 1082 "Else" "noBreak"
              $ 1083 "PSE_T≔get_random_pose(pose_ref=CAM_Pose, mode='rotation', range_max=[10,10,0])"
              global PSE_T=get_random_pose(pose_ref=CAM_Pose, mode="rotation", range_max=[10,10,0])
              $ 1084 "CAM_LM_Refined≔ True "
              global CAM_LM_Refined=  True
            end
            $ 1085 "If get_inverse_kin_has_solution(pose_trans(FRM_Reference, PSE_T))"
            if (get_inverse_kin_has_solution( pose_trans (FRM_Reference, PSE_T))):
              $ 1086 "Comment"
              # Comment
              $ 1087 "PSE_T" "breakAfter"
              set_tcp(p[0.0,0.0,0.161,3.1415,0.0,0.0])
              movel(pose_trans(FRM_Reference, PSE_T), a=0.03, v=0.05)
            else:
              $ 1088 "Else" "noBreak"
              $ 1089 "'If random pose is out of reach, set the initial cam pose'"
              # 'If random pose is out of reach, set the initial cam pose'
              $ 1090 "PSE_T≔CAM_Pose"
              global PSE_T=CAM_Pose
            end
          end
        end
        $ 1091 "Wait: 2.0"
        sleep(2.0)
        $ 1092 "trigger"
        $ 1093 "If ITM_ID≟1 and JIG≟7"
        if (ITM_ID == 1  and  JIG == 7):
          # begin: URCap Program Node
          #   Source: SensoPart VISOR Robotic, 2.0.6, SensoPart Industriesensorik GmbH
          #   Type: VISOR Trigger
          $ 1094 "# 1 VISOR Trigger"
          visor_changeJob(1, "Landmark_INVITE_2", 6000)
          visor_trigger(1, 6000, "arm")
          # end: URCap Program Node
        else:
          $ 1095 "ElseIf ITM_ID≟5 and JIG≟7"
          if (ITM_ID == 5  and  JIG == 7):
            # begin: URCap Program Node
            #   Source: SensoPart VISOR Robotic, 2.0.6, SensoPart Industriesensorik GmbH
            #   Type: VISOR Trigger
            $ 1096 "# 1 VISOR Trigger"
            visor_changeJob(1, "Landmark_INVITE_2", 6000)
            visor_trigger(1, 6000, "arm")
            # end: URCap Program Node
          else:
            $ 1097 "ElseIf ITM_ID≟13 and JIG≟7"
            if (ITM_ID == 13  and  JIG == 7):
              # begin: URCap Program Node
              #   Source: SensoPart VISOR Robotic, 2.0.6, SensoPart Industriesensorik GmbH
              #   Type: VISOR Trigger
              $ 1098 "# 1 VISOR Trigger"
              visor_changeJob(1, "Landmark_INVITE_2", 6000)
              visor_trigger(1, 6000, "arm")
              # end: URCap Program Node
            else:
              $ 1099 "ElseIf ITM_ID≟1 and JIG≟15"
              if (ITM_ID == 1 and JIG == 15):
                # begin: URCap Program Node
                #   Source: SensoPart VISOR Robotic, 2.0.6, SensoPart Industriesensorik GmbH
                #   Type: VISOR Trigger
                $ 1100 "# 1 VISOR Trigger"
                visor_changeJob(1, "Aztec_no_dot_pick", 6000)
                visor_trigger(1, 6000, "arm")
                # end: URCap Program Node
              else:
                $ 1101 "ElseIf ITM_ID≟1 and JIG≟21"
                if (ITM_ID == 1 and JIG == 21):
                  # begin: URCap Program Node
                  #   Source: SensoPart VISOR Robotic, 2.0.6, SensoPart Industriesensorik GmbH
                  #   Type: VISOR Trigger
                  $ 1102 "# 1 VISOR Trigger"
                  visor_changeJob(1, "PoTS", 6000)
                  visor_trigger(1, 6000, "arm")
                  # end: URCap Program Node
                else:
                  $ 1103 "ElseIf ITM_ID≟1 and JIG≟17"
                  if (ITM_ID == 1 and JIG == 17):
                    # begin: URCap Program Node
                    #   Source: SensoPart VISOR Robotic, 2.0.6, SensoPart Industriesensorik GmbH
                    #   Type: VISOR Trigger
                    $ 1104 "# 1 VISOR Trigger"
                    visor_changeJob(1, "Weigh_target", 6000)
                    visor_trigger(1, 6000, "arm")
                    # end: URCap Program Node
                  end
                end
              end
            end
          end
        end
        $ 1108 "TM_3D_Found≔visor_partsFound(1)"
        global TM_3D_Found= visor_partsFound (1)
        $ 1110 "If TM_3D_Found>0"
        if (TM_3D_Found>0):
          $ 1111 "CAM_LM_Detected≔ True "
          global CAM_LM_Detected=  True
          $ 1112 "CAM_Captures≔0"
          global CAM_Captures=0
        else:
          $ 1113 "Else" "noBreak"
          $ 1114 "CAM_LM_Detected≔ False "
          global CAM_LM_Detected=  False
          $ 1115 "CAM_Captures≔CAM_Captures+1"
          global CAM_Captures=CAM_Captures+1
        end
        $ 1120 "result"
        $ 1121 "If CAM_LM_Detected"
        if (CAM_LM_Detected):
          $ 1122 "If (CAM_LM_Refinmnt and CAM_LM_Refined) or  not CAM_LM_Refinmnt"
          if ((CAM_LM_Refinmnt  and  CAM_LM_Refined)  or    not  CAM_LM_Refinmnt):
            $ 1180 "If ITM_ID≟1 and JIG≟7"
            if (ITM_ID == 1  and  JIG == 7):
              $ 1181 "CAM_LM_SSRack≔visor_getPose3d(1, 0)"
              global CAM_LM_SSRack= visor_getPose3d (1, 0)
            else:
              $ 1182 "ElseIf ITM_ID≟5 and JIG≟7"
              if (ITM_ID == 5  and  JIG == 7):
                $ 1183 "CAM_LM_SSRack≔visor_getPose3d(1, 0)"
                global CAM_LM_SSRack= visor_getPose3d (1, 0)
              else:
                $ 1186 "ElseIf ITM_ID≟1 and JIG≟15"
                if (ITM_ID == 1 and JIG == 15):
                  $ 1187 "CAM_LM_cont≔visor_getPose3d(1, 0)"
                  global CAM_LM_cont= visor_getPose3d (1, 0)
                  $ 1188 "Trigger≔get_actual_tcp_pose()"
                  global Trigger= get_actual_tcp_pose ()
                else:
                  $ 1189 "ElseIf ITM_ID≟1 and JIG≟21"
                  if (ITM_ID == 1 and JIG == 21):
                    $ 1190 "CAM_LM_cont≔visor_getPose3d(1, 0)"
                    global CAM_LM_cont= visor_getPose3d (1, 0)
                    $ 1191 "Trigger≔get_actual_tcp_pose()"
                    global Trigger= get_actual_tcp_pose ()
                  else:
                    $ 1192 "ElseIf ITM_ID≟1 and JIG≟17"
                    if (ITM_ID == 1 and JIG == 17):
                      $ 1193 "CAM_LM_cont≔visor_getPose3d(1, 0)"
                      global CAM_LM_cont= visor_getPose3d (1, 0)
                      $ 1194 "Trigger≔get_actual_tcp_pose()"
                      global Trigger= get_actual_tcp_pose ()
                    end
                  end
                end
              end
            end
            $ 1195 "CAM_Done≔ True "
            global CAM_Done=  True
          end
        else:
          $ 1196 "ElseIf  not CAM_LM_Detected and CAM_Captures<CAM_PRM_Retries"
          if (  not  CAM_LM_Detected  and  CAM_Captures<CAM_PRM_Retries):
            $ 1197 "CAM_LM_Refined≔ False "
            global CAM_LM_Refined=  False
          else:
            $ 1198 "ElseIf CAM_Captures≥CAM_PRM_Retries"
            if (CAM_Captures >= CAM_PRM_Retries):
              $ 1199 "CAM_Done≔ True "
              global CAM_Done=  True
              $ 1200 "Error"
              $ 1201 "set_error(ERROR_NO_LANDMARK)"
              set_error(ERROR_NO_LANDMARK)
            end
          end
        end
      end
    elif (151 == switch_1):
      $ 1202 "Case 151"
      $ 1203 "Detect (SensoPart)"
      $ 1204 "go to capture pose"
      $ 1205 "FRM_Reference≔FRM_Cap_SSRack"
      global FRM_Reference=FRM_Cap_SSRack
      $ 1206 "PSE_T≔p[0,0,-0.00,0,0,0]"
      global PSE_T=p[0,0,-0.00,0,0,0]
      $ 1207 "do_transition(pose_trans(FRM_Reference, PSE_T), keep_rxry=False)"
      do_transition( pose_trans (FRM_Reference, PSE_T), keep_rxry=False)
      $ 1208 "JNT_Q≔get_actual_joint_positions()"
      global JNT_Q= get_actual_joint_positions ()
      $ 1209 "JNT_Q≔[JNT_Q[0], JNT_Q[1], JNT_Q[2], JNT_Q[3], JNT_Q[4], 0]"
      global JNT_Q=[JNT_Q[0], JNT_Q[1], JNT_Q[2], JNT_Q[3], JNT_Q[4], 0]
      $ 1210 "Set"
      set_tcp(p[0.0,0.0,0.161,3.1415,0.0,0.0])
      $ 1211 "movej(get_inverse_kin(pose_trans(FRM_Reference, PSE_T), qnear=JNT_Q))"
      movej(get_inverse_kin( pose_trans (FRM_Reference, PSE_T), qnear=JNT_Q))
      $ 1212 "CAM_Pose≔pose_trans(pose_inv(FRM_Reference), get_actual_tcp_pose())"
      global CAM_Pose= pose_trans ( pose_inv (FRM_Reference),  get_actual_tcp_pose ())
      $ 1213 "Loop  not CAM_Done and  not ERROR.FLAG and  not CMD_Stop"
      while (  not  CAM_Done  and    not  ERROR.FLAG  and    not  CMD_Stop):
        $ 1214 "If  not OBJ_Detected and CAM_Captures>0"
        if (  not  OBJ_Detected  and  CAM_Captures>0):
          $ 1215 "MoveL"
          $ 1216 "If FRM_Reference≟p[0,0,0,0,0,0]"
          if (FRM_Reference == p[0,0,0,0,0,0]):
            $ 1218 "PSE_T≔get_random_pose(pose_ref=CAM_Pose, mode='rotation', range_max=[15,15,0])"
            global PSE_T=get_random_pose(pose_ref=CAM_Pose, mode="rotation", range_max=[15,15,0])
          else:
            $ 1219 "Else" "noBreak"
            $ 1220 "PSE_T≔get_random_pose(pose_ref=CAM_Pose, mode='rotation', range_max=[10,10,0])"
            global PSE_T=get_random_pose(pose_ref=CAM_Pose, mode="rotation", range_max=[10,10,0])
          end
          $ 1221 "If get_inverse_kin_has_solution(pose_trans(FRM_Reference, PSE_T))"
          if (get_inverse_kin_has_solution( pose_trans (FRM_Reference, PSE_T))):
            $ 1222 "PSE_T" "breakAfter"
            set_tcp(p[0.0,0.0,0.161,3.1415,0.0,0.0])
            movel(pose_trans(FRM_Reference, PSE_T), a=0.03, v=0.05)
          else:
            $ 1223 "Else" "noBreak"
            $ 1224 "'If random pose is out of reach, set the initial cam pose'"
            # 'If random pose is out of reach, set the initial cam pose'
            $ 1225 "PSE_T≔CAM_Pose"
            global PSE_T=CAM_Pose
            $ 1226 "PSE_T" "breakAfter"
            set_tcp(p[0.0,0.0,0.161,3.1415,0.0,0.0])
            movel(pose_trans(FRM_Reference, PSE_T), a=0.03, v=0.05)
          end
        end
        $ 1227 "Wait: 0.5"
        sleep(0.5)
        $ 1228 "Set"
        set_tcp(p[0.0,0.0,0.161,3.1415,0.0,0.0])
        # begin: URCap Program Node
        #   Source: SensoPart VISOR Robotic, 2.0.6, SensoPart Industriesensorik GmbH
        #   Type: VISOR Trigger
        $ 1229 "# 1 VISOR Trigger"
        visor_changeJob(1, "Object Detection Single", 6000)
        visor_trigger(1, 6000, "arm")
        # end: URCap Program Node
        $ 1230 "If visor_isResponseOk(1)"
        if ( visor_isResponseOk (1)):
          $ 1231 "CAM_CNT_Obj≔visor_partsFound(1)"
          global CAM_CNT_Obj= visor_partsFound (1)
          $ 1232 "CAM_OBJ_Pose≔visor_getPose3d(1, 0)"
          global CAM_OBJ_Pose= visor_getPose3d (1, 0)
          $ 1233 "If CAM_CNT_Obj>0"
          if (CAM_CNT_Obj>0):
            $ 1234 "CAM_OBJ_Color≔visor_getAdditionalData(1, 0)"
            global CAM_OBJ_Color= visor_getAdditionalData (1, 0)
            $ 1235 "CAM_DetectScore≔to_num(visor_getAdditionalData(1, 1))/1000"
            global CAM_DetectScore=to_num( visor_getAdditionalData (1, 1))/1000
            $ 1236 "OBJ_Detected≔ True "
            global OBJ_Detected=  True
          end
        else:
          $ 1237 "Else" "noBreak"
          $ 1238 "CAM_Captures≔CAM_Captures+1"
          global CAM_Captures=CAM_Captures+1
        end
        $ 1239 "If OBJ_Detected"
        if (OBJ_Detected):
          $ 1240 "Get object data"
          $ 1241 "PRC_CntDetect≔0"
          global PRC_CntDetect=0
          $ 1242 "Loop PRC_CntDetect<CAM_CNT_Obj"
          while (PRC_CntDetect<CAM_CNT_Obj):
            $ 1243 "get object and jig number"
            $ 1244 "If ITM_ID≟1 and JIG≟7"
            if (ITM_ID == 1  and  JIG == 7):
              $ 1245 "FRM_Reference≔FRM_Cap_SSRack"
              global FRM_Reference=FRM_Cap_SSRack
            else:
              $ 1246 "ElseIf ITM_ID≟5 and JIG≟7"
              if (ITM_ID == 5  and  JIG == 7):
                $ 1247 "FRM_Reference≔uLM_Cap_SSRack"
                global FRM_Reference=uLM_Cap_SSRack
              end
            end
            $ 1250 "PSE_T≔pose_trans(pose_inv(FRM_Reference), CAM_OBJ_Pose)"
            global PSE_T= pose_trans ( pose_inv (FRM_Reference), CAM_OBJ_Pose)
            $ 1251 "CAM_Result.append(get_pattern_counter(PSE_T, 'X', pattern=[10, 5], patternsize=[0.181, 0.081]))"
            CAM_Result.append(get_pattern_counter(PSE_T, "X", pattern=[10, 5], patternsize=[0.181, 0.081]))
            $ 1252 "PRC_CntDetect≔PRC_CntDetect+1"
            global PRC_CntDetect=PRC_CntDetect+1
          end
          $ 1253 "CAM_Done≔ True "
          global CAM_Done=  True
        else:
          $ 1254 "ElseIf CAM_Captures≥CAM_PRM_Retries"
          if (CAM_Captures >= CAM_PRM_Retries):
            $ 1255 "CAM_Done≔ True "
            global CAM_Done=  True
          else:
            $ 1256 "Else" "noBreak"
            $ 1257 "CAM_Captures≔CAM_Captures+1"
            global CAM_Captures=CAM_Captures+1
          end
        end
      end
    end
    $ 1258 "'=========='"
    # '=========='
    $ 1259 "PostSettings"
    $ 1260 "FRM_Reference≔p[0,0,0,0,0,0]"
    global FRM_Reference=p[0,0,0,0,0,0]
    $ 1261 "Set"
    set_tcp(p[0.0,0.0,0.161,3.1415,0.0,0.0])
    $ 1262 "CAM_Pose≔p[0,0,0,0,0,0]"
    global CAM_Pose=p[0,0,0,0,0,0]
    $ 1263 "Action≔0"
    global Action=0
    $ 1264 "Action_Info≔''"
    global Action_Info=""
  end
  def Sub_AMR_MiR_V3():
    $ 1265 "Sub_AMR_MiR_V3" "noBreak"
    $ 1266 "PreSettings"
    $ 1267 "AMR_TargetList≔[1,2,3,4,5,21,22,23,24,31,32,33,34,35,36,37,38,41]"
    global AMR_TargetList=[1,2,3,4,5,21,22,23,24,31,32,33,34,35,36,37,38,41]
    $ 1268 "AMR_Done≔ False "
    global AMR_Done=  False
    $ 1269 "AMR_PosActual≔T2O_Current_Pos"
    global AMR_PosActual=modbus_get_signal_status("T2O_Current_Pos")
    $ 1270 "AMR_Attemps≔T2O_Nav_Attemps"
    global AMR_Attemps=modbus_get_signal_status("T2O_Nav_Attemps")
    $ 1271 "AMR_Battery≔MiR_Battery_Lvl"
    global AMR_Battery=modbus_get_signal_status("MiR_Battery_Lvl")
    $ 1272 "AMR_Charging≔(T2O_Charging≟1)"
    global AMR_Charging=(modbus_get_signal_status("T2O_Charging") == 1)
    $ 1273 "AMR_Position≔struct(position_identifier=T2O_Current_Pos, x1=MiR_Position_X1, x2=MiR_Position_X2, y1=MiR_Position_Y1, y2=MiR_Position_Y2, theta1=MiR_Theta_1, theta2=MiR_Theta_2) "
    global AMR_Position=struct(position_identifier=modbus_get_signal_status("T2O_Current_Pos"), x1=modbus_get_signal_status("MiR_Position_X1"), x2=modbus_get_signal_status("MiR_Position_X2"), y1=modbus_get_signal_status("MiR_Position_Y1"), y2=modbus_get_signal_status("MiR_Position_Y2"), theta1=modbus_get_signal_status("MiR_Theta_1"), theta2=modbus_get_signal_status("MiR_Theta_2"))
    $ 1274 "If MiR_Mode≠7"
    if (modbus_get_signal_status("MiR_Mode") != 7):
      $ 1275 "Error"
      $ 1276 "set_error(ERROR_AMR_WRONG_MODE)"
      set_error(ERROR_AMR_WRONG_MODE)
      $ 1277 "AMR_Done≔ True "
      global AMR_Done=  True
    end
    $ 1278 "'=========='"
    # '=========='
    $ 1279 "Switch STATE"
    switch_1 = STATE
    $ 1280 "Case 1"
    if (1 == switch_1):
      $ 1281 "stopping"
      $ 1282 "If T2O_Done≟1 and O2T_Acknowledge≟0"
      if (modbus_get_signal_status("T2O_Done") == 1  and  modbus_get_signal_status("O2T_Acknowledge") == 0):
        $ 1283 "Set O2T_Acknowledge=1"
        modbus_set_output_register("O2T_Acknowledge", 1)
      end
      $ 1284 "Set MiR_CMD_Stop=On"
      modbus_set_output_signal("MiR_CMD_Stop", True)
      $ 1285 "AMR_Position.position_identifier = 0"
      AMR_Position.position_identifier = 0
      $ 1286 "AMR_Done≔ True "
      global AMR_Done=  True
    elif (2 == switch_1):
      $ 1287 "Case 2"
      $ 1288 "stopped"
      $ 1289 "If MiR_State≠3 and MiR_State≠5"
      if (modbus_get_signal_status("MiR_State") != 3  and  modbus_get_signal_status("MiR_State") != 5):
        $ 1290 "Set MiR_CMD_Stop=Off"
        modbus_set_output_signal("MiR_CMD_Stop", False)
      end
    elif (3 == switch_1):
      $ 1291 "Case 3"
      $ 1292 "resetting"
      $ 1293 "Set O2T_Mis_Main=Off"
      modbus_set_output_signal("O2T_Mis_Main", False)
      $ 1294 "Set O2T_Mis_Charge=Off"
      modbus_set_output_signal("O2T_Mis_Charge", False)
      $ 1295 "If MiR_Mis_Queue>0"
      if (modbus_get_signal_status("MiR_Mis_Queue")>0):
        $ 1296 "Set MiR_CMD_Clear_Q=On"
        modbus_set_output_signal("MiR_CMD_Clear_Q", True)
        $ 1297 "Wait MiR_Mis_Queue≟0"
        while (not(modbus_get_signal_status("MiR_Mis_Queue") == 0)):
          sync()
        end
        $ 1298 "Set MiR_CMD_Clear_Q=Off"
        modbus_set_output_signal("MiR_CMD_Clear_Q", False)
      end
      $ 1299 "If MiR_Error_ID≠0"
      if (modbus_get_signal_status("MiR_Error_ID") != 0):
        $ 1300 "Set MiR_CMD_Clear_E=On"
        modbus_set_output_signal("MiR_CMD_Clear_E", True)
        $ 1301 "Wait MiR_Error_ID≟0"
        while (not(modbus_get_signal_status("MiR_Error_ID") == 0)):
          sync()
        end
        $ 1302 "Set MiR_CMD_Clear_E=Off"
        modbus_set_output_signal("MiR_CMD_Clear_E", False)
      end
      $ 1303 "Set O2T_Action=0"
      modbus_set_output_register("O2T_Action", 0)
      $ 1304 "Set O2T_Acknowledge=0"
      modbus_set_output_register("O2T_Acknowledge", 0)
      $ 1305 "Set O2T_Target_Pos=0"
      modbus_set_output_register("O2T_Target_Pos", 0)
      $ 1306 "Set O2T_Footprint=0"
      modbus_set_output_register("O2T_Footprint", 0)
      $ 1307 "Set O2T_ProtectOff=0"
      modbus_set_output_register("O2T_ProtectOff", 0)
      $ 1308 "Set O2T_Dock=0"
      modbus_set_output_register("O2T_Dock", 0)
      $ 1309 "AMR_Attemps≔0"
      global AMR_Attemps=0
      $ 1310 "AMR_PosTarget≔0"
      global AMR_PosTarget=0
      $ 1311 "AMR_Step≔0"
      global AMR_Step=0
      $ 1312 "AMR_AtTarget≔ False "
      global AMR_AtTarget=  False
      $ 1313 "If MiR_State≟4 or MiR_State≟3 or MiR_State≟10"
      if (modbus_get_signal_status("MiR_State") == 4  or  modbus_get_signal_status("MiR_State") == 3  or  modbus_get_signal_status("MiR_State") == 10):
        $ 1314 "AMR_Done≔ True "
        global AMR_Done=  True
      end
    elif (5 == switch_1):
      $ 1315 "Case 5"
      $ 1316 "starting"
      $ 1317 "If MiR_State≟4"
      if (modbus_get_signal_status("MiR_State") == 4):
        $ 1318 "Set MiR_CMD_Start=On"
        modbus_set_output_signal("MiR_CMD_Start", True)
        $ 1319 "Wait MiR_State≠4"
        while (not(modbus_get_signal_status("MiR_State") != 4)):
          sync()
        end
        $ 1320 "Set MiR_CMD_Start=Off"
        modbus_set_output_signal("MiR_CMD_Start", False)
        $ 1321 "AMR_Done≔ True "
        global AMR_Done=  True
      else:
        $ 1322 "ElseIf MiR_State≟10"
        if (modbus_get_signal_status("MiR_State") == 10):
          $ 1323 "'MiR in protective stop. Wait'"
          # 'MiR in protective stop. Wait'
          $ 1324 "AMR_Done≔ True "
          global AMR_Done=  True
        else:
          $ 1325 "ElseIf MiR_State≟3"
          if (modbus_get_signal_status("MiR_State") == 3):
            $ 1326 "AMR_Done≔ True "
            global AMR_Done=  True
          end
        end
      end
    elif (6 == switch_1):
      $ 1327 "Case 6"
      $ 1328 "execute"
      $ 1329 "AMR_AtTarget≔(AMR_PosActual≟AMR_PosTarget)"
      global AMR_AtTarget=(AMR_PosActual == AMR_PosTarget)
      $ 1330 "Switch AMR_Step"
      switch_2 = AMR_Step
      $ 1331 "Case 0"
      if (0 == switch_2):
        $ 1332 "If  not AMR_AtTarget"
        if (  not  AMR_AtTarget):
          $ 1333 "AMR_Step≔1"
          global AMR_Step=1
        else:
          $ 1334 "Else" "noBreak"
          $ 1335 "AMR_Done≔ True "
          global AMR_Done=  True
        end
      elif (1 == switch_2):
        $ 1336 "Case 1"
        $ 1337 "general Settings"
        $ 1338 "Set O2T_Acknowledge=0"
        modbus_set_output_register("O2T_Acknowledge", 0)
        $ 1339 "check for error"
        $ 1340 "If OBJ_Picked and MiR_State≟10"
        if (OBJ_Picked  and  modbus_get_signal_status("MiR_State") == 10):
          $ 1341 "Error"
          $ 1342 "set_error(ERROR_ROBOT_ARM_NOT_IN_HOME_POSE)"
          set_error(ERROR_ROBOT_ARM_NOT_IN_HOME_POSE)
          $ 1343 "Action≔0"
          global Action=0
        else:
          $ 1344 "ElseIf  not found_in_list(AMR_PosTarget, AMR_TargetList)"
          if (  not  found_in_list(AMR_PosTarget, AMR_TargetList)):
            $ 1345 "Error"
            $ 1346 "set_error(ERROR_UNKNOWN_POSE)"
            set_error(ERROR_UNKNOWN_POSE)
            $ 1347 "Action≔0"
            global Action=0
          end
        end
        $ 1348 "If MiR_State≟3"
        if (modbus_get_signal_status("MiR_State") == 3):
          $ 1349 "Set MiR_CMD_Start=Off"
          modbus_set_output_signal("MiR_CMD_Start", False)
          $ 1350 "Switch Action"
          switch_3 = Action
          $ 1351 "Case 51"
          if (51 == switch_3):
            $ 1352 "Charge"
            $ 1353 "'trigger the charging mission'"
            # 'trigger the charging mission'
            $ 1354 "'target pos is predefined'"
            # 'target pos is predefined'
            $ 1355 "Set O2T_Footprint=0"
            modbus_set_output_register("O2T_Footprint", 0)
            $ 1356 "Set O2T_Action=1"
            modbus_set_output_register("O2T_Action", 1)
            $ 1357 "If MiR_Mis_Queue≟0"
            if (modbus_get_signal_status("MiR_Mis_Queue") == 0):
              $ 1358 "Set O2T_Mis_Charge=On"
              modbus_set_output_signal("O2T_Mis_Charge", True)
              $ 1359 "Wait MiR_Mis_Queue≥1"
              while (not(modbus_get_signal_status("MiR_Mis_Queue") >= 1)):
                sync()
              end
              $ 1360 "Set O2T_Mis_Charge=Off"
              modbus_set_output_signal("O2T_Mis_Charge", False)
            end
          elif (52 == switch_3):
            $ 1361 "Case 52"
            $ 1362 "Navigate"
            $ 1363 "'trigger the standard missoin'"
            # 'trigger the standard missoin'
            $ 1364 "Set O2T_Footprint=AMR_FootprintID"
            modbus_set_output_register("O2T_Footprint", AMR_FootprintID)
            $ 1365 "Set O2T_Target_Pos=AMR_PosTarget"
            modbus_set_output_register("O2T_Target_Pos", AMR_PosTarget)
            $ 1366 "Set O2T_Action=2"
            modbus_set_output_register("O2T_Action", 2)
            $ 1367 "If MiR_Mis_Queue≟0"
            if (modbus_get_signal_status("MiR_Mis_Queue") == 0):
              $ 1368 "Set O2T_Mis_Main=On"
              modbus_set_output_signal("O2T_Mis_Main", True)
              $ 1369 "Wait MiR_Mis_Queue≥1"
              while (not(modbus_get_signal_status("MiR_Mis_Queue") >= 1)):
                sync()
              end
              $ 1370 "Set O2T_Mis_Main=Off"
              modbus_set_output_signal("O2T_Mis_Main", False)
            end
          end
        else:
          $ 1371 "ElseIf MiR_State≟4"
          if (modbus_get_signal_status("MiR_State") == 4):
            $ 1372 "Set MiR_CMD_Start=On"
            modbus_set_output_signal("MiR_CMD_Start", True)
          else:
            $ 1373 "ElseIf MiR_State≟5"
            if (modbus_get_signal_status("MiR_State") == 5):
              $ 1374 "AMR_Step≔2"
              global AMR_Step=2
            else:
              $ 1375 "ElseIf MiR_State≟10"
              if (modbus_get_signal_status("MiR_State") == 10):
                $ 1376 "'AMR still in safeguard stop'"
                # 'AMR still in safeguard stop'
              end
            end
          end
        end
      elif (2 == switch_2):
        $ 1377 "Case 2"
        $ 1378 "acknowledge handshake"
        $ 1379 "If T2O_Done≟1 and O2T_Acknowledge≟0"
        if (modbus_get_signal_status("T2O_Done") == 1  and  modbus_get_signal_status("O2T_Acknowledge") == 0):
          $ 1380 "Set O2T_Acknowledge=1"
          modbus_set_output_register("O2T_Acknowledge", 1)
        else:
          $ 1381 "ElseIf T2O_Done≟0 and O2T_Acknowledge≟1"
          if (modbus_get_signal_status("T2O_Done") == 0  and  modbus_get_signal_status("O2T_Acknowledge") == 1):
            $ 1382 "Set O2T_Acknowledge=0"
            modbus_set_output_register("O2T_Acknowledge", 0)
            $ 1383 "AMR_AtTarget≔(AMR_PosActual≟AMR_PosTarget)"
            global AMR_AtTarget=(AMR_PosActual == AMR_PosTarget)
            $ 1384 "AMR_Done≔ True "
            global AMR_Done=  True
          end
        end
      end
      $ 1385 "translate errors"
      $ 1386 "If AMR_Done"
      if (AMR_Done):
        $ 1387 "Switch T2O_Error_ID"
        switch_2 = modbus_get_signal_status("T2O_Error_ID")
        $ 1388 "Case 2003"
        if (2003 == switch_2):
          $ 1389 "error"
          $ 1390 "set_error(ERROR_NOT_DOCKED)"
          set_error(ERROR_NOT_DOCKED)
        elif (2007 == switch_2):
          $ 1391 "Case 2007"
          $ 1392 "error"
          $ 1393 "set_error(ERROR_NOT_REACHABLE_TARGET)"
          set_error(ERROR_NOT_REACHABLE_TARGET)
        elif (2008 == switch_2):
          $ 1394 "Case 2008"
          $ 1395 "error"
          $ 1396 "set_error(ERROR_CHARGING_NOT_STARTED)"
          set_error(ERROR_CHARGING_NOT_STARTED)
        end
      end
    elif (7 == switch_1):
      $ 1397 "Case 7"
      $ 1398 "completing"
      $ 1399 "If MiR_Mis_Queue>0"
      if (modbus_get_signal_status("MiR_Mis_Queue")>0):
        $ 1400 "Set MiR_CMD_Abort=On"
        modbus_set_output_signal("MiR_CMD_Abort", True)
        $ 1401 "Wait MiR_Mis_Queue≟0"
        while (not(modbus_get_signal_status("MiR_Mis_Queue") == 0)):
          sync()
        end
        $ 1402 "Set MiR_CMD_Abort=Off"
        modbus_set_output_signal("MiR_CMD_Abort", False)
      end
      $ 1403 "If MiR_State≟3 or MiR_State≟10"
      if (modbus_get_signal_status("MiR_State") == 3  or  modbus_get_signal_status("MiR_State") == 10):
        $ 1404 "AMR_Done≔ True "
        global AMR_Done=  True
      end
    elif (9 == switch_1):
      $ 1405 "Case 9"
      $ 1406 "holding"
      $ 1407 "Set MiR_CMD_Abort=On"
      modbus_set_output_signal("MiR_CMD_Abort", True)
      $ 1408 "If MiR_State≟3 or MiR_State≟10"
      if (modbus_get_signal_status("MiR_State") == 3  or  modbus_get_signal_status("MiR_State") == 10):
        $ 1409 "Set MiR_CMD_Abort=Off"
        modbus_set_output_signal("MiR_CMD_Abort", False)
        $ 1410 "AMR_Done≔ True "
        global AMR_Done=  True
      end
    elif (11 == switch_1):
      $ 1411 "Case 11"
      $ 1412 "unholding"
      $ 1413 "Set MiR_CMD_Start=On"
      modbus_set_output_signal("MiR_CMD_Start", True)
      $ 1414 "If MiR_State≠4"
      if (modbus_get_signal_status("MiR_State") != 4):
        $ 1415 "Set MiR_CMD_Start=Off"
        modbus_set_output_signal("MiR_CMD_Start", False)
        $ 1416 "AMR_Step≔0"
        global AMR_Step=0
        $ 1417 "AMR_Done≔ True "
        global AMR_Done=  True
      end
    elif (12 == switch_1):
      $ 1418 "Case 12"
      $ 1419 "suspending"
      $ 1420 "'none'"
      # 'none'
    elif (14 == switch_1):
      $ 1421 "Case 14"
      $ 1422 "unsuspending"
      $ 1423 "'none'"
      # 'none'
    elif (15 == switch_1):
      $ 1424 "Case 15"
      $ 1425 "aborting"
      $ 1426 "Set MiR_CMD_Abort=On"
      modbus_set_output_signal("MiR_CMD_Abort", True)
      $ 1427 "Wait MiR_State≟3"
      while (not(modbus_get_signal_status("MiR_State") == 3)):
        sync()
      end
      $ 1428 "Set MiR_CMD_Abort=Off"
      modbus_set_output_signal("MiR_CMD_Abort", False)
    elif (17 == switch_1):
      $ 1429 "Case 17"
      $ 1430 "clearing"
      $ 1431 "If MiR_Error_ID≠0"
      if (modbus_get_signal_status("MiR_Error_ID") != 0):
        $ 1432 "Set MiR_CMD_Clear_E=On"
        modbus_set_output_signal("MiR_CMD_Clear_E", True)
        $ 1433 "Wait MiR_Error_ID≟0"
        while (not(modbus_get_signal_status("MiR_Error_ID") == 0)):
          sync()
        end
        $ 1434 "Set MiR_CMD_Clear_E=Off"
        modbus_set_output_signal("MiR_CMD_Clear_E", False)
      end
      $ 1435 "If MiR_Error_ID≟0"
      if (modbus_get_signal_status("MiR_Error_ID") == 0):
        $ 1436 "AMR_Done≔ True "
        global AMR_Done=  True
      end
    end
    $ 1437 "'=========='"
    # '=========='
    $ 1438 "PostSettings"
    $ 1439 "AMR_Position≔struct(position_identifier=T2O_Current_Pos, x1=MiR_Position_X1, x2=MiR_Position_X2, y1=MiR_Position_Y1, y2=MiR_Position_Y2, theta1=MiR_Theta_1, theta2=MiR_Theta_2) "
    global AMR_Position=struct(position_identifier=modbus_get_signal_status("T2O_Current_Pos"), x1=modbus_get_signal_status("MiR_Position_X1"), x2=modbus_get_signal_status("MiR_Position_X2"), y1=modbus_get_signal_status("MiR_Position_Y1"), y2=modbus_get_signal_status("MiR_Position_Y2"), theta1=modbus_get_signal_status("MiR_Theta_1"), theta2=modbus_get_signal_status("MiR_Theta_2"))
  end
  def Sub_Action_V4():
    $ 1440 "Sub_Action_V4" "noBreak"
    $ 1441 "PreSettings"
    $ 1442 "init poses"
    $ 1443 "PSE_A≔p[0,0,0,0,0,0]"
    global PSE_A=p[0,0,0,0,0,0]
    $ 1444 "PSE_A_H≔p[0,0,0,0,0,0]"
    global PSE_A_H=p[0,0,0,0,0,0]
    $ 1445 "PSE_T≔p[0,0,0,0,0,0]"
    global PSE_T=p[0,0,0,0,0,0]
    $ 1446 "PSE_T_H≔p[0,0,0,0,0,0]"
    global PSE_T_H=p[0,0,0,0,0,0]
    $ 1447 "PSE_G≔p[0,0,0,0,0,0]"
    global PSE_G=p[0,0,0,0,0,0]
    $ 1448 "PSE_G_H≔p[0,0,0,0,0,0]"
    global PSE_G_H=p[0,0,0,0,0,0]
    $ 1449 "PSE_R≔p[0,0,0,0,0,0]"
    global PSE_R=p[0,0,0,0,0,0]
    $ 1450 "PSE_R_H≔p[0,0,0,0,0,0]"
    global PSE_R_H=p[0,0,0,0,0,0]
    $ 1451 "JNT_Q≔[0,0,0,0,0,0]"
    global JNT_Q=[0,0,0,0,0,0]
    $ 1452 "JNT_S≔[0,0,0,0,0,0]"
    global JNT_S=[0,0,0,0,0,0]
    $ 1453 "Gripping parameters"
    $ 1454 "OBJ = find_object_by_type(OBJs, OBJ_Type)"
    OBJ = find_object_by_type(OBJs, OBJ_Type)
    $ 1455 "GRP_Open_Pos≔OBJ.dimension.diameter * 1000 + 6"
    global GRP_Open_Pos=OBJ.dimension.diameter * 1000 + 6
    $ 1456 "GRP_Offset≔OBJ.gripper_offset"
    global GRP_Offset=OBJ.gripper_offset
    $ 1457 "rq_set_force_norm(50)"
     rq_set_force_norm (50)
    $ 1458 "rq_set_speed_norm(50)"
     rq_set_speed_norm (50)
    $ 1459 "Switch ITM_ID"
    switch_1 = ITM_ID
    $ 1460 "Case 1"
    if (1 == switch_1):
      $ 1461 "uML"
      $ 1462 "JIG2 = find_object_by_type(JIGs, JIG)"
      JIG2 = find_object_by_type(JIGs, JIG)
      $ 1463 "JIG_Offset≔JIG2.jig_offset"
      global JIG_Offset=JIG2.jig_offset
      $ 1464 "Switch JIG"
      switch_2 = JIG
      $ 1465 "Case 1"
      if (1 == switch_2):
        $ 1466 "3FG"
        $ 1467 "define poses"
        $ 1468 "FRM_Reference≔ULM_3FG"
        global FRM_Reference=ULM_3FG
        $ 1469 "JNT_Q≔JNT_HOME"
        global JNT_Q=JNT_HOME
        $ 1470 "PSE_T≔pose_trans(GRP_Offset, JIG_Offset)"
        global PSE_T= pose_trans (GRP_Offset, JIG_Offset)
        $ 1471 "PSE_A≔pose_trans(PSE_T, p[0,0,0.100,0,0,0])"
        global PSE_A= pose_trans (PSE_T, p[0,0,0.100,0,0,0])
        $ 1472 "PSE_R≔pose_add(PSE_T, p[0,0,0.100,0,0,0])"
        global PSE_R= pose_add (PSE_T, p[0,0,0.100,0,0,0])
      elif (2 == switch_2):
        $ 1473 "Case 2"
        $ 1474 "Input"
        $ 1475 "'CHANGE THE REFERENCE TO THE FRAME TO MOVE IN'"
        # 'CHANGE THE REFERENCE TO THE FRAME TO MOVE IN'
        $ 1476 "define poses"
        $ 1477 "FRM_Reference≔ULM_Input"
        global FRM_Reference=ULM_Input
        $ 1478 "PSE_T≔pose_trans(pose_trans(get_pattern_pos_rectangle(OBJ_Nbr, 'X', [10,5], patternsize=[0.181,0.081]), GRP_Offset), JIG_Offset)"
        global PSE_T= pose_trans ( pose_trans (get_pattern_pos_rectangle(OBJ_Nbr, "X", [10,5], patternsize=[0.181,0.081]), GRP_Offset), JIG_Offset)
        $ 1479 "If Action≟1"
        if (Action == 1):
          $ 1480 "PSE_R≔pose_add(PSE_T, p[0,0,0.200,0,0,0])"
          global PSE_R= pose_add (PSE_T, p[0,0,0.200,0,0,0])
          $ 1481 "PSE_A≔pose_add(PSE_T, p[0,0,0.100,0,0,0])"
          global PSE_A= pose_add (PSE_T, p[0,0,0.100,0,0,0])
        else:
          $ 1482 "ElseIf Action≟2"
          if (Action == 2):
            $ 1483 "PSE_R≔pose_add(PSE_T, p[0,0,0.100,0,0,0])"
            global PSE_R= pose_add (PSE_T, p[0,0,0.100,0,0,0])
            $ 1484 "PSE_A≔pose_add(PSE_T, p[0,0,0.200,0,0,0])"
            global PSE_A= pose_add (PSE_T, p[0,0,0.200,0,0,0])
          end
        end
      elif (3 == switch_2):
        $ 1485 "Case 3"
        $ 1486 "Output"
        $ 1487 "'CHANGE THE REFERENCE TO THE FRAME TO MOVE IN'"
        # 'CHANGE THE REFERENCE TO THE FRAME TO MOVE IN'
        $ 1488 "define poses"
        $ 1489 "FRM_Reference≔ULM_Output"
        global FRM_Reference=ULM_Output
        $ 1490 "PSE_T≔pose_trans(pose_trans(get_pattern_pos_rectangle(OBJ_Nbr, 'X', [10,5], patternsize=[0.181,0.081]), GRP_Offset), JIG_Offset)"
        global PSE_T= pose_trans ( pose_trans (get_pattern_pos_rectangle(OBJ_Nbr, "X", [10,5], patternsize=[0.181,0.081]), GRP_Offset), JIG_Offset)
        $ 1492 "If Action≟1"
        if (Action == 1):
          $ 1493 "PSE_R≔pose_add(PSE_T, p[0,0,0.200,0,0,0])"
          global PSE_R= pose_add (PSE_T, p[0,0,0.200,0,0,0])
          $ 1494 "PSE_A≔pose_add(PSE_T, p[0,0,0.100,0,0,0])"
          global PSE_A= pose_add (PSE_T, p[0,0,0.100,0,0,0])
        else:
          $ 1495 "ElseIf Action≟2"
          if (Action == 2):
            $ 1496 "PSE_R≔pose_add(PSE_T, p[0,0,0.100,0,0,0])"
            global PSE_R= pose_add (PSE_T, p[0,0,0.100,0,0,0])
            $ 1497 "PSE_A≔pose_add(PSE_T, p[0,0,0.200,0,0,0])"
            global PSE_A= pose_add (PSE_T, p[0,0,0.200,0,0,0])
          end
        end
      elif (4 == switch_2):
        $ 1498 "Case 4"
        $ 1499 "jig centrifuge racks"
        $ 1500 "define poses"
        $ 1501 "FRM_Reference≔ULM_Cent_Racks"
        global FRM_Reference=ULM_Cent_Racks
        $ 1502 "PSE_T≔get_pattern_pos_rectangle(JIG_Slot, 'X', [4,1], patternsize=[0.291,0])"
        global PSE_T=get_pattern_pos_rectangle(JIG_Slot, "X", [4,1], patternsize=[0.291,0])
        $ 1503 "If OBJ_Nbr≠0"
        if (OBJ_Nbr != 0):
          $ 1504 "PSE_T≔pose_trans(pose_trans(PSE_T, get_pattern_pos_rectangle(OBJ_Nbr, 'X', [3,3], patternsize=[0.060,0.060])),p[-0.030, -0.030,0,0,0,3.927])"
          global PSE_T= pose_trans ( pose_trans (PSE_T, get_pattern_pos_rectangle(OBJ_Nbr, "X", [3,3], patternsize=[0.060,0.060])),p[-0.030, -0.030,0,0,0,3.927])
        end
        $ 1505 "PSE_T≔pose_trans(PSE_T, GRP_Offset)"
        global PSE_T= pose_trans (PSE_T, GRP_Offset)
        $ 1506 "If Action≟1"
        if (Action == 1):
          $ 1507 "PSE_R≔pose_add(PSE_T, p[0,0,0.200,0,0,0])"
          global PSE_R= pose_add (PSE_T, p[0,0,0.200,0,0,0])
          $ 1508 "PSE_A≔pose_add(PSE_T, p[0,0,0.100,0,0,0])"
          global PSE_A= pose_add (PSE_T, p[0,0,0.100,0,0,0])
        else:
          $ 1509 "ElseIf Action≟2"
          if (Action == 2):
            $ 1510 "PSE_R≔pose_add(PSE_T, p[0,0,0.100,0,0,0])"
            global PSE_R= pose_add (PSE_T, p[0,0,0.100,0,0,0])
            $ 1511 "PSE_A≔pose_add(PSE_T, p[0,0,0.200,0,0,0])"
            global PSE_A= pose_add (PSE_T, p[0,0,0.200,0,0,0])
          end
        end
      elif (6 == switch_2):
        $ 1512 "Case 6"
        $ 1513 "Caps bin"
        $ 1514 "define poses"
        $ 1515 "'Drop cap'"
        # 'Drop cap'
        $ 1516 "FRM_Reference=ULM_Cap_Bin"
        FRM_Reference=ULM_Cap_Bin
        $ 1517 "PSE_T≔pose_RPY2RotVec(p[0,0,0,0,0,0])"
        global PSE_T=pose_RPY2RotVec(p[0,0,0,0,0,0])
        $ 1518 "PSE_T_H≔pose_add(PSE_T, p[0,0,-0.011,0,0,0])"
        global PSE_T_H= pose_add (PSE_T, p[0,0,-0.011,0,0,0])
        $ 1519 "PSE_A≔pose_trans(PSE_T, p[0,0,0.1,0,0,0])"
        global PSE_A= pose_trans (PSE_T, p[0,0,0.1,0,0,0])
        $ 1520 "PSE_R_H≔pose_add(PSE_T, p[0,0,0.100,0,0,0])"
        global PSE_R_H= pose_add (PSE_T, p[0,0,0.100,0,0,0])
        $ 1521 "PSE_R≔pose_add(PSE_T, p[0,0,0.100,0,0,0])"
        global PSE_R= pose_add (PSE_T, p[0,0,0.100,0,0,0])
      elif (7 == switch_2):
        $ 1522 "Case 7"
      elif (8 == switch_2):
        $ 1547 "Case 8"
        $ 1548 "NoK"
        $ 1549 "define poses"
        $ 1550 "'NoK'"
        # 'NoK'
        $ 1551 "FRM_Reference=ULM_NoK"
        FRM_Reference=ULM_NoK
        $ 1552 "PSE_T≔pose_RPY2RotVec(p[0,0,0,0,0,0])"
        global PSE_T=pose_RPY2RotVec(p[0,0,0,0,0,0])
        $ 1553 "PSE_A≔pose_trans(PSE_T, p[0,0,0.1,0,0,0])"
        global PSE_A= pose_trans (PSE_T, p[0,0,0.1,0,0,0])
        $ 1554 "PSE_R≔pose_add(PSE_T, p[0,0,0.100,0,0,0])"
        global PSE_R= pose_add (PSE_T, p[0,0,0.100,0,0,0])
      elif (9 == switch_2):
        $ 1555 "Case 9"
      elif (10 == switch_2):
        $ 1563 "Case 10"
      elif (11 == switch_2):
        $ 1571 "Case 11"
      elif (12 == switch_2):
        $ 1579 "Case 12"
      end
    elif (2 == switch_1):
      $ 1587 "Case 2"
      $ 1588 "Centrifuge"
      $ 1589 "'CHANGE THE REFERENCE TO THE FRAME TO MOVE IN'"
      # 'CHANGE THE REFERENCE TO THE FRAME TO MOVE IN'
      $ 1590 "define poses"
      $ 1591 "FRM_Reference≔FRM_Centrifuge"
      global FRM_Reference=FRM_Centrifuge
      $ 1592 "PSE_T≔GRP_Offset"
      global PSE_T=GRP_Offset
      $ 1593 "If Action≟8"
      if (Action == 8):
        $ 1594 "PSE_R≔pose_add(PSE_T, p[0,0,0.250,0,0,0])"
        global PSE_R= pose_add (PSE_T, p[0,0,0.250,0,0,0])
        $ 1595 "PSE_A≔pose_add(PSE_T, p[0,0,0.150,0,0,0])"
        global PSE_A= pose_add (PSE_T, p[0,0,0.150,0,0,0])
      else:
        $ 1596 "ElseIf Action≟7"
        if (Action == 7):
          $ 1597 "PSE_R≔pose_add(PSE_T, p[0,0,0.150,0,0,0])"
          global PSE_R= pose_add (PSE_T, p[0,0,0.150,0,0,0])
          $ 1598 "PSE_A≔pose_add(PSE_T, p[0,0,0.250,0,0,0])"
          global PSE_A= pose_add (PSE_T, p[0,0,0.250,0,0,0])
        end
      end
    elif (3 == switch_1):
      $ 1599 "Case 3"
      $ 1600 "Output"
      $ 1601 "'CHANGE THE REFERENCE TO THE FRAME TO MOVE IN'"
      # 'CHANGE THE REFERENCE TO THE FRAME TO MOVE IN'
      $ 1602 "define poses"
      $ 1603 "FRM_Reference≔Base_const"
      global FRM_Reference=p[0.0,0.0,0.0,0.0,0.0,0.0]
      $ 1604 "PSE_T≔p[0,0,0,0,0,0]"
      global PSE_T=p[0,0,0,0,0,0]
      $ 1605 "PSE_A≔pose_add(PSE_T, p[0,0,0.150,0,0,0])"
      global PSE_A= pose_add (PSE_T, p[0,0,0.150,0,0,0])
      $ 1606 "PSE_R≔pose_add(PSE_T, p[0,0,0.100,0,0,0])"
      global PSE_R= pose_add (PSE_T, p[0,0,0.100,0,0,0])
    elif (5 == switch_1):
      $ 1607 "Case 5"
      $ 1608 "Sarstedt Pickup Table"
      $ 1609 "'CHANGE THE REFERENCE TO THE FRAME TO MOVE IN'"
      # 'CHANGE THE REFERENCE TO THE FRAME TO MOVE IN'
      $ 1610 "Switch JIG"
      switch_2 = JIG
      $ 1611 "Case 7"
      if (7 == switch_2):
        $ 1624 "Sarstedt"
        $ 1625 "'CHANGE THE REFERENCE TO THE FRAME TO MOVE IN'"
        # 'CHANGE THE REFERENCE TO THE FRAME TO MOVE IN'
        $ 1631 "If TASK.ID≟10"
        if (TASK.ID == 10):
          $ 1632 "Frame & Position Params"
          $ 1633 "FRM_Reference = CAM_LM_SSRack"
          FRM_Reference = CAM_LM_SSRack
          $ 1634 "PSE_T≔uLM_SS_PickPlc"
          global PSE_T=uLM_SS_PickPlc
          $ 1635 "PSE_A≔pose_trans(PSE_T, p[0,0,0.1,0,0,0])"
          global PSE_A= pose_trans (PSE_T, p[0,0,0.1,0,0,0])
          $ 1636 "PSE_R≔pose_add(PSE_T, p[0,0,0.1,0,0,0])"
          global PSE_R= pose_add (PSE_T, p[0,0,0.1,0,0,0])
        end
      end
    elif (13 == switch_1):
      $ 1643 "Case 13"
      $ 1644 "Sarstedt Pickup Table"
      $ 1645 "'CHANGE THE REFERENCE TO THE FRAME TO MOVE IN'"
      # 'CHANGE THE REFERENCE TO THE FRAME TO MOVE IN'
      $ 1646 "Switch JIG"
      switch_2 = JIG
      $ 1647 "Case 7"
      if (7 == switch_2):
        $ 1660 "Bottle"
        $ 1661 "'CHANGE THE REFERENCE TO THE FRAME TO MOVE IN'"
        # 'CHANGE THE REFERENCE TO THE FRAME TO MOVE IN'
        $ 1667 "If TASK.ID≟43"
        if (TASK.ID == 43):
          $ 1668 "Frame & Position Params"
          $ 1670 "PSE_T≔uLM_SS_PickPlc"
          global PSE_T=uLM_SS_PickPlc
          $ 1671 "PSE_A≔pose_trans(PSE_T, p[0,0,0.1,0,0,0])"
          global PSE_A= pose_trans (PSE_T, p[0,0,0.1,0,0,0])
          $ 1672 "PSE_R≔pose_add(PSE_T, p[0,0,0.1,0,0,0])"
          global PSE_R= pose_add (PSE_T, p[0,0,0.1,0,0,0])
        end
      end
    end
    $ 1679 "Additional check"
    $ 1680 "If  not is_reachable(FRM_Reference,[PSE_A,PSE_A_H,PSE_T,PSE_T_H,PSE_R,PSE_R_H])"
    if (  not  is_reachable(FRM_Reference,[PSE_A,PSE_A_H,PSE_T,PSE_T_H,PSE_R,PSE_R_H])):
      $ 1681 "Error"
      $ 1682 "set_error(ERROR_POSE_NOT_REACHABLE)"
      set_error(ERROR_POSE_NOT_REACHABLE)
      $ 1683 "Action≔0"
      global Action=0
    end
    $ 1684 "'=========='"
    # '=========='
    $ 1685 "Switch Action"
    switch_1 = Action
    $ 1686 "Case 1"
    if (1 == switch_1):
      $ 1687 "Pick"
      $ 1688 "Action_Info≔'pick object'"
      global Action_Info="pick object"
      $ 1689 "do_transition(pose_trans(FRM_Reference, PSE_T), keep_rxry=OBJ_Picked)"
      do_transition( pose_trans (FRM_Reference, PSE_T), keep_rxry=OBJ_Picked)
      $ 1690 "EOAT"
      $ 1691 "If  not OBJ_Picked"
      if (  not  OBJ_Picked):
        $ 1692 "rq_move_and_wait_mm(GRP_Open_Pos)"
         rq_move_and_wait_mm (GRP_Open_Pos)
      end
      $ 1693 "If PSE_A_H≠PSE_Z"
      if (PSE_A_H != PSE_Z):
        $ 1694 "If JNT_Q≠JNT_Z"
        if (JNT_Q != JNT_Z):
          $ 1695 "movej(get_inverse_kin(pose_trans(FRM_Reference, PSE_A_H), qnear=JNT_Q), r=0.050)"
          movej(get_inverse_kin( pose_trans (FRM_Reference, PSE_A_H), qnear=JNT_Q), r=0.050)
        else:
          $ 1696 "Else" "noBreak"
          $ 1697 "movej(pose_trans(FRM_Reference, PSE_A_H), r=0.050)"
          movej( pose_trans (FRM_Reference, PSE_A_H), r=0.050)
        end
      end
      $ 1698 "If PSE_A≠PSE_Z"
      if (PSE_A != PSE_Z):
        $ 1699 "If JNT_Q≠JNT_Z"
        if (JNT_Q != JNT_Z):
          $ 1700 "movej(get_inverse_kin(pose_trans(FRM_Reference, PSE_A), qnear=JNT_Q), r=0.020)"
          movej(get_inverse_kin( pose_trans (FRM_Reference, PSE_A), qnear=JNT_Q), r=0.020)
        else:
          $ 1701 "Else" "noBreak"
          $ 1702 "movej(pose_trans(FRM_Reference, PSE_A), r=0.020)"
          movej( pose_trans (FRM_Reference, PSE_A), r=0.020)
        end
      end
      $ 1703 "MoveL"
      $ 1704 "If PSE_T_H≠PSE_Z"
      if (PSE_T_H != PSE_Z):
        $ 1705 "PSE_T_H" "breakAfter"
        movel(pose_trans(FRM_Reference, PSE_T_H), a=0.5, v=0.4, r=0.01)
      end
      $ 1706 "PSE_T" "breakAfter"
      movel(pose_trans(FRM_Reference, PSE_T), a=0.08, v=0.12)
      $ 1707 "EOAT"
      $ 1708 "rq_set_force_norm(50)"
       rq_set_force_norm (50)
      $ 1709 "rq_close_and_wait()"
       rq_close_and_wait ()
      $ 1710 "OBJ_Picked≔rq_is_object_detected()"
      global OBJ_Picked= rq_is_object_detected ()
      $ 1711 "If  not OBJ_Picked"
      if (  not  OBJ_Picked):
        $ 1712 "set_error(ERROR_NO_OBJECT_TO_PICK)"
        set_error(ERROR_NO_OBJECT_TO_PICK)
      end
      $ 1713 "EXTT"
      $ 1714 "Switch JIG"
      switch_2 = JIG
      $ 1715 "Case 1"
      if (1 == switch_2):
        $ 1716 "3FG"
        $ 1717 "If OBJ_Picked"
        if (OBJ_Picked):
          $ 1718 "Set GRP_3F_Open=On"
          set_standard_digital_out(5, True)
        end
      end
      $ 1719 "If PSE_R_H≠PSE_Z"
      if (PSE_R_H != PSE_Z):
        $ 1720 "PSE_R" "breakAfter"
        movel(pose_trans(FRM_Reference, PSE_R), a=0.5, v=0.4, r=0.01)
        $ 1721 "PSE_R_H" "breakAfter"
        movel(pose_trans(FRM_Reference, PSE_R_H), a=0.5, v=0.4)
      else:
        $ 1722 "Else" "noBreak"
        $ 1723 "PSE_R" "breakAfter"
        movel(pose_trans(FRM_Reference, PSE_R), a=0.5, v=0.4)
      end
    elif (2 == switch_1):
      $ 1724 "Case 2"
      $ 1725 "Place"
      $ 1726 "Action_Info≔'place object'"
      global Action_Info="place object"
      $ 1727 "do_transition(pose_trans(FRM_Reference, PSE_T), keep_rxry=OBJ_Picked)"
      do_transition( pose_trans (FRM_Reference, PSE_T), keep_rxry=OBJ_Picked)
      $ 1728 "EXTT"
      $ 1729 "Switch JIG"
      switch_2 = JIG
      $ 1730 "Case 1"
      if (1 == switch_2):
        $ 1731 "3FG"
        $ 1732 "If OBJ_Picked"
        if (OBJ_Picked):
          $ 1733 "Set GRP_3F_Open=On"
          set_standard_digital_out(5, True)
        end
      end
      $ 1734 "If PSE_A_H≠PSE_Z"
      if (PSE_A_H != PSE_Z):
        $ 1735 "If JNT_Q≠JNT_Z"
        if (JNT_Q != JNT_Z):
          $ 1736 "movej(get_inverse_kin(pose_trans(FRM_Reference, PSE_A_H), qnear=JNT_Q), r=0.050)"
          movej(get_inverse_kin( pose_trans (FRM_Reference, PSE_A_H), qnear=JNT_Q), r=0.050)
        else:
          $ 1737 "Else" "noBreak"
          $ 1738 "movej(pose_trans(FRM_Reference, PSE_A_H), r=0.050)"
          movej( pose_trans (FRM_Reference, PSE_A_H), r=0.050)
        end
      end
      $ 1739 "If PSE_A≠PSE_Z"
      if (PSE_A != PSE_Z):
        $ 1740 "If JNT_Q≠JNT_Z"
        if (JNT_Q != JNT_Z):
          $ 1741 "movej(get_inverse_kin(pose_trans(FRM_Reference, PSE_A), qnear=JNT_Q), r=0.020)"
          movej(get_inverse_kin( pose_trans (FRM_Reference, PSE_A), qnear=JNT_Q), r=0.020)
        else:
          $ 1742 "Else" "noBreak"
          $ 1743 "movej(pose_trans(FRM_Reference, PSE_A), r=0.020)"
          movej( pose_trans (FRM_Reference, PSE_A), r=0.020)
        end
      end
      $ 1744 "MoveL"
      $ 1745 "If PSE_T_H≠PSE_Z"
      if (PSE_T_H != PSE_Z):
        $ 1746 "PSE_T_H" "breakAfter"
        movel(pose_trans(FRM_Reference, PSE_T_H), a=0.5, v=0.4, r=0.01)
      end
      $ 1747 "PSE_T" "breakAfter"
      global move_thread_flag_1747=0
      thread move_thread_1747():
        enter_critical
        move_thread_flag_1747 = 1
        movel(pose_trans(FRM_Reference, PSE_T), a=0.05, v=0.09)
        move_thread_flag_1747 = 2
        exit_critical
      end
      move_thread_flag_1747 = 0
      move_thread_han_1747 = run move_thread_1747()
      while (True):
        local targetTcpDirection=get_target_tcp_speed()
        local stepsToRetract=tool_contact(direction=targetTcpDirection)
        if (stepsToRetract > 0):
          kill move_thread_han_1747
          stopl(0.5)
          $ 1748 "Until (tool_contact_detection)"
          break
        end
        sleep(1.0E-10)
        if (move_thread_flag_1747 > 1):
          join move_thread_han_1747
          break
        end
        sync()
      end
      $ 1749 "Force"
      sleep(0.02)
      zero_ftsensor()
      force_mode(FRM_Reference, [1, 1, 1, 0, 0, 0], [0.0, 0.0, 0.0, 0.0, 0.0, 0.0], 2, [0.1, 0.1, 0.01, 0.3490658503988659, 0.3490658503988659, 0.3490658503988659])
      $ 1750 "PSE_T" "noBreak"
      movel(pose_trans(FRM_Reference, PSE_T), a=0.04, v=0.07)
      end_force_mode()
      stopl(5.0)
      $ 1751 "EXTT"
      $ 1752 "Switch JIG"
      switch_2 = JIG
      $ 1753 "Case 1"
      if (1 == switch_2):
        $ 1754 "3FG"
        $ 1755 "If OBJ_Picked"
        if (OBJ_Picked):
          $ 1756 "Set GRP_3F_Open=Off"
          set_standard_digital_out(5, False)
          $ 1757 "Wait: 0.2"
          sleep(0.2)
        end
      end
      $ 1758 "EOAT"
      $ 1759 "rq_move_and_wait_mm(GRP_Open_Pos)"
       rq_move_and_wait_mm (GRP_Open_Pos)
      $ 1760 "OBJ_Picked≔rq_is_object_detected()"
      global OBJ_Picked= rq_is_object_detected ()
      $ 1761 "If PSE_R_H≠PSE_Z"
      if (PSE_R_H != PSE_Z):
        $ 1762 "PSE_R" "breakAfter"
        movel(pose_trans(FRM_Reference, PSE_R), a=0.5, v=0.4, r=0.01)
        $ 1763 "PSE_R_H" "breakAfter"
        movel(pose_trans(FRM_Reference, PSE_R_H), a=0.5, v=0.4)
      else:
        $ 1764 "Else" "noBreak"
        $ 1765 "PSE_R" "breakAfter"
        movel(pose_trans(FRM_Reference, PSE_R), a=0.5, v=0.4)
      end
    elif (3 == switch_1):
      $ 1766 "Case 3"
      $ 1767 "Push"
      $ 1768 "Action_Info≔'push'"
      global Action_Info="push"
    elif (4 == switch_1):
      $ 1769 "Case 4"
      $ 1770 "Pull"
      $ 1771 "Action_Info≔'pull'"
      global Action_Info="pull"
    elif (6 == switch_1):
      $ 1774 "Case 6"
      $ 1775 "Drop the cap"
      $ 1776 "If JNT_A≠[0,0,0,0,0,0]"
      if (JNT_A != [0,0,0,0,0,0]):
        $ 1777 "MoveJ"
        $ 1778 "JNT_A" "breakAfter"
        movej(JNT_A, a=1.3962634015954636, v=1.7453292519943295, r=0.02)
      else:
        $ 1779 "Else" "noBreak"
        $ 1780 "MoveJ"
        $ 1781 "PSE_A" "breakAfter"
        movej(pose_trans(FRM_Reference, PSE_A), a=1.3962634015954636, v=1.7453292519943295, r=0.02)
      end
      $ 1782 "MoveL"
      $ 1783 "PSE_T" "breakAfter"
      movel(pose_trans(FRM_Reference, PSE_T), a=0.05, v=0.09)
      $ 1784 "'ADD OPEN GRIPPER'"
      # 'ADD OPEN GRIPPER'
      # begin: URCap Program Node
      #   Source: Robotiq_Grippers, 3.17.0.105337, Robotiq Inc.
      #   Type: Gripper
      $ 1785 "Gripper Move10mm (1)"
      if not(gripper_connected[0]):
        popup("Gripper 1 must be connected to run this program.", "No connection", False, True, True)
      end
      if not(rq_is_gripper_activated("1")):
        popup("Gripper 1 is not activated. Go to Installation tab > Gripper to activate it and run the program again.", "Not activated", False, True, True)
      end
      rq_set_pos_spd_for(201, 0, 28, "1")
      rq_wait_pos_spe_for_request(201, 0, 28, "1")
      rq_go_to("1")
      rq_wait("1")
      # end: URCap Program Node
      $ 1786 "PSE_T_H" "breakAfter"
      movel(pose_trans(FRM_Reference, PSE_T_H), a=0.05, v=0.09)
      # begin: URCap Program Node
      #   Source: Robotiq_Grippers, 3.17.0.105337, Robotiq Inc.
      #   Type: Gripper
      $ 1787 "Gripper Move40mm (1)"
      if not(gripper_connected[0]):
        popup("Gripper 1 must be connected to run this program.", "No connection", False, True, True)
      end
      if not(rq_is_gripper_activated("1")):
        popup("Gripper 1 is not activated. Go to Installation tab > Gripper to activate it and run the program again.", "Not activated", False, True, True)
      end
      rq_set_pos_spd_for(63, 0, 28, "1")
      rq_wait_pos_spe_for_request(63, 0, 28, "1")
      rq_go_to("1")
      rq_wait("1")
      # end: URCap Program Node
      $ 1788 "PSE_R" "breakAfter"
      movel(pose_trans(FRM_Reference, PSE_R), a=0.5, v=0.4)
    elif (7 == switch_1):
      $ 1789 "Case 7"
      $ 1790 "Load"
      $ 1791 "Action_Info≔'load object'"
      global Action_Info="load object"
      $ 1792 "do_transition(pose_trans(FRM_Reference, PSE_T), keep_rxry=OBJ_Picked)"
      do_transition( pose_trans (FRM_Reference, PSE_T), keep_rxry=OBJ_Picked)
      $ 1793 "If PSE_A_H≠PSE_Z"
      if (PSE_A_H != PSE_Z):
        $ 1794 "If JNT_Q≠JNT_Z"
        if (JNT_Q != JNT_Z):
          $ 1795 "movej(get_inverse_kin(pose_trans(FRM_Reference, PSE_A_H), qnear=JNT_Q), r=0.050)"
          movej(get_inverse_kin( pose_trans (FRM_Reference, PSE_A_H), qnear=JNT_Q), r=0.050)
        else:
          $ 1796 "Else" "noBreak"
          $ 1797 "movej(pose_trans(FRM_Reference, PSE_A_H), r=0.050)"
          movej( pose_trans (FRM_Reference, PSE_A_H), r=0.050)
        end
      end
      $ 1798 "If PSE_A≠PSE_Z"
      if (PSE_A != PSE_Z):
        $ 1799 "If JNT_Q≠JNT_Z"
        if (JNT_Q != JNT_Z):
          $ 1800 "movej(get_inverse_kin(pose_trans(FRM_Reference, PSE_A), qnear=JNT_Q), r=0.020)"
          movej(get_inverse_kin( pose_trans (FRM_Reference, PSE_A), qnear=JNT_Q), r=0.020)
        else:
          $ 1801 "Else" "noBreak"
          $ 1802 "movej(pose_trans(FRM_Reference, PSE_A), r=0.020)"
          movej( pose_trans (FRM_Reference, PSE_A), r=0.020)
        end
      end
      $ 1803 "MoveL"
      $ 1804 "If PSE_T_H≠PSE_Z"
      if (PSE_T_H != PSE_Z):
        $ 1805 "PSE_T_H" "breakAfter"
        movel(pose_trans(FRM_Reference, PSE_T_H), a=0.5, v=0.4, r=0.01)
      end
      $ 1806 "PSE_T" "breakAfter"
      global move_thread_flag_1806=0
      thread move_thread_1806():
        enter_critical
        move_thread_flag_1806 = 1
        movel(pose_trans(FRM_Reference, PSE_T), a=0.05, v=0.09)
        move_thread_flag_1806 = 2
        exit_critical
      end
      move_thread_flag_1806 = 0
      move_thread_han_1806 = run move_thread_1806()
      while (True):
        local targetTcpDirection=get_target_tcp_speed()
        local stepsToRetract=tool_contact(direction=targetTcpDirection)
        if (stepsToRetract > 0):
          kill move_thread_han_1806
          stopl(0.5)
          $ 1807 "Until (tool_contact_detection)"
          break
        end
        sleep(1.0E-10)
        if (move_thread_flag_1806 > 1):
          join move_thread_han_1806
          break
        end
        sync()
      end
      $ 1808 "Force"
      sleep(0.02)
      zero_ftsensor()
      force_mode(FRM_Reference, [0, 1, 1, 0, 0, 1], [0.0, 0.0, 0.0, 0.0, 0.0, 0.0], 2, [0.1, 0.05, 0.02, 0.3490658503988659, 0.3490658503988659, 3.141592653589793])
      $ 1809 "PSE_T" "noBreak"
      movel(pose_trans(FRM_Reference, PSE_T), a=0.04, v=0.07)
      end_force_mode()
      stopl(5.0)
      $ 1810 "EOAT"
      $ 1811 "rq_move_and_wait_mm(GRP_Open_Pos)"
       rq_move_and_wait_mm (GRP_Open_Pos)
      $ 1812 "OBJ_Picked≔rq_is_object_detected()"
      global OBJ_Picked= rq_is_object_detected ()
      $ 1813 "If PSE_R_H≠PSE_Z"
      if (PSE_R_H != PSE_Z):
        $ 1814 "PSE_R" "breakAfter"
        movel(pose_trans(FRM_Reference, PSE_R), a=0.5, v=0.4, r=0.01)
        $ 1815 "PSE_R_H" "breakAfter"
        movel(pose_trans(FRM_Reference, PSE_R_H), a=0.5, v=0.4)
      else:
        $ 1816 "Else" "noBreak"
        $ 1817 "PSE_R" "breakAfter"
        movel(pose_trans(FRM_Reference, PSE_R), a=0.5, v=0.4)
      end
    elif (8 == switch_1):
      $ 1818 "Case 8"
      $ 1819 "Unload"
      $ 1820 "Action_Info≔'pick object'"
      global Action_Info="pick object"
      $ 1821 "do_transition(pose_trans(FRM_Reference, PSE_T), keep_rxry=OBJ_Picked)"
      do_transition( pose_trans (FRM_Reference, PSE_T), keep_rxry=OBJ_Picked)
      $ 1822 "EOAT"
      $ 1823 "If  not OBJ_Picked"
      if (  not  OBJ_Picked):
        $ 1824 "rq_move_and_wait_mm(GRP_Open_Pos)"
         rq_move_and_wait_mm (GRP_Open_Pos)
      end
      $ 1825 "If PSE_A_H≠PSE_Z"
      if (PSE_A_H != PSE_Z):
        $ 1826 "If JNT_Q≠JNT_Z"
        if (JNT_Q != JNT_Z):
          $ 1827 "movej(get_inverse_kin(pose_trans(FRM_Reference, PSE_A_H), qnear=JNT_Q), r=0.050)"
          movej(get_inverse_kin( pose_trans (FRM_Reference, PSE_A_H), qnear=JNT_Q), r=0.050)
        else:
          $ 1828 "Else" "noBreak"
          $ 1829 "movej(pose_trans(FRM_Reference, PSE_A_H), r=0.050)"
          movej( pose_trans (FRM_Reference, PSE_A_H), r=0.050)
        end
      end
      $ 1830 "If PSE_A≠PSE_Z"
      if (PSE_A != PSE_Z):
        $ 1831 "If JNT_Q≠JNT_Z"
        if (JNT_Q != JNT_Z):
          $ 1832 "movej(get_inverse_kin(pose_trans(FRM_Reference, PSE_A), qnear=JNT_Q), r=0.020)"
          movej(get_inverse_kin( pose_trans (FRM_Reference, PSE_A), qnear=JNT_Q), r=0.020)
        else:
          $ 1833 "Else" "noBreak"
          $ 1834 "movej(pose_trans(FRM_Reference, PSE_A), r=0.020)"
          movej( pose_trans (FRM_Reference, PSE_A), r=0.020)
        end
      end
      $ 1835 "MoveL"
      $ 1836 "If PSE_T_H≠PSE_Z"
      if (PSE_T_H != PSE_Z):
        $ 1837 "PSE_T_H" "breakAfter"
        movel(pose_trans(FRM_Reference, PSE_T_H), a=0.5, v=0.4, r=0.01)
      end
      $ 1838 "PSE_T" "breakAfter"
      movel(pose_trans(FRM_Reference, PSE_T), a=0.08, v=0.12)
      $ 1839 "Force"
      sleep(0.02)
      zero_ftsensor()
      force_mode(FRM_Reference, [1, 1, 0, 0, 0, 0], [0.0, 0.0, 0.0, 0.0, 0.0, 0.0], 2, [0.05, 0.05, 0.1, 0.3490658503988659, 0.3490658503988659, 0.3490658503988659])
      $ 1840 "EOAT" "noBreak"
      $ 1841 "rq_set_force_norm(50)" "noBreak"
       rq_set_force_norm (50)
      $ 1842 "rq_close_and_wait()" "noBreak"
       rq_close_and_wait ()
      $ 1843 "OBJ_Picked≔rq_is_object_detected()" "noBreak"
      global OBJ_Picked= rq_is_object_detected ()
      $ 1844 "If  not OBJ_Picked" "noBreak"
      if (  not  OBJ_Picked):
        $ 1845 "set_error(ERROR_NO_OBJECT_TO_PICK)" "noBreak"
        set_error(ERROR_NO_OBJECT_TO_PICK)
      end
      $ 1846 "If PSE_R_H≠PSE_Z" "noBreak"
      if (PSE_R_H != PSE_Z):
        $ 1847 "PSE_R" "noBreak"
        movel(pose_trans(FRM_Reference, PSE_R), a=0.5, v=0.4, r=0.01)
        $ 1848 "PSE_R_H" "noBreak"
        movel(pose_trans(FRM_Reference, PSE_R_H), a=0.5, v=0.4)
      else:
        $ 1849 "Else" "noBreak"
        $ 1850 "PSE_R" "noBreak"
        movel(pose_trans(FRM_Reference, PSE_R), a=0.5, v=0.4)
      end
      end_force_mode()
      stopl(5.0)
    elif (11 == switch_1):
      $ 1851 "Case 11"
    elif (12 == switch_1):
      $ 1888 "Case 12"
      $ 1889 "Decap"
      $ 1890 "Action_Info≔'decapping'"
      global Action_Info="decapping"
      $ 1891 "Set GRP_3F_Enable=On"
      set_standard_digital_out(4, True)
      $ 1892 "Set GRP_3F_Decap=On"
      set_standard_digital_out(3, True)
      $ 1893 "Force"
      sleep(0.02)
      zero_ftsensor()
      force_mode(tool_pose(), [0, 0, 1, 0, 0, 0], [0.0, 0.0, 5.0, 0.0, 0.0, 0.0], 2, [0.1, 0.1, 0.15, 0.3490658503988659, 0.3490658503988659, 0.3490658503988659])
      $ 1894 "check_decapping(offset=0.015, timeout=5, abort=CMD_Hold)" "noBreak"
      check_decapping(offset=0.015, timeout=5, abort=CMD_Hold)
      end_force_mode()
      stopl(5.0)
      $ 1895 "Set GRP_3F_Decap=Off"
      set_standard_digital_out(3, False)
      $ 1896 "Set GRP_3F_Enable=Off"
      set_standard_digital_out(4, False)
      $ 1897 "MoveL"
      $ 1898 "PSE_R" "breakAfter"
      movel(pose_trans(FRM_Reference, PSE_R), a=0.8, v=0.15)
    elif (13 == switch_1):
      $ 1899 "Case 13"
      $ 1900 "TMR_Barcode: Reset"
      TMR_Barcode = 0
      $ 1901 "Read"
      $ 1902 "TMR_Barcode: Start"
      TMR_Barcode_is_counting = True
      $ 1903 "If TMR_Barcode<PRM_TO_Read_BC"
      global thread_flag_1903=0
      thread Thread_if_1903():
        $ 1904 "KeyenceTrigger"
        $ 1905 "Set OClearResult=HI:Pulse 0.2"
        thread SinglePulse4():
          write_output_boolean_register(2, True)
          sleep(0.2)
          write_output_boolean_register(2, False)
        end
        singlePulse4 = run SinglePulse4()
        $ 1906 "Wait: 0.5"
        sleep(0.5)
        $ 1907 "Set OTriggerBarcode=Off"
        write_output_boolean_register(1, False)
        $ 1908 "Wait: 0.5"
        sleep(0.5)
        $ 1909 "Set OTriggerBarcode=On"
        write_output_boolean_register(1, True)
        $ 1910 "Wait: 0.5"
        sleep(0.5)
        $ 1911 "Preorient"
        $ 1912 "TMR_Barcode: Reset"
        TMR_Barcode = 0
        $ 1913 "If ICmdExctd"
        if (read_input_boolean_register(12)):
          $ 1914 "Set GRP_3F_Decap=On"
          set_standard_digital_out(3, True)
          $ 1915 "Set GRP_3F_Enable=On"
          set_standard_digital_out(4, True)
          $ 1916 "Loop ICmdExctd"
          while (read_input_boolean_register(12)):
            $ 1917 "KeyenceTrigger"
            $ 1918 "Set OClearResult=HI:Pulse 0.1"
            thread SinglePulse5():
              write_output_boolean_register(2, True)
              sleep(0.1)
              write_output_boolean_register(2, False)
            end
            singlePulse5 = run SinglePulse5()
            $ 1919 "Wait: 0.3"
            sleep(0.3)
            $ 1920 "Set OTriggerBarcode=Off"
            write_output_boolean_register(1, False)
            $ 1921 "Wait: 0.3"
            sleep(0.3)
            $ 1922 "Set OTriggerBarcode=On"
            write_output_boolean_register(1, True)
            $ 1923 "Wait: 0.1"
            sleep(0.1)
          end
        end
        $ 1924 "If  not ICmdExctd"
        if (  not  read_input_boolean_register(12)):
          $ 1925 "Set GRP_3F_Decap=On"
          set_standard_digital_out(3, True)
          $ 1926 "Set GRP_3F_Enable=On"
          set_standard_digital_out(4, True)
          $ 1927 "Wait ICmdExctd=HI"
          while (read_input_boolean_register(12) == False):
            sync()
          end
        end
        $ 1928 "Set GRP_3F_Decap=Off"
        set_standard_digital_out(3, False)
        $ 1929 "Set GRP_3F_Enable=Off"
        set_standard_digital_out(4, False)
        $ 1930 "OBJ_Brc_OK≔ True "
        global OBJ_Brc_OK=  True
        thread_flag_1903 = 1
      end
      if (TMR_Barcode<PRM_TO_Read_BC):
        global thread_handler_1903=run Thread_if_1903()
        while (thread_flag_1903 == 0):
          if not(TMR_Barcode<PRM_TO_Read_BC):
            kill thread_handler_1903
            thread_flag_1903 = 2
          else:
            sync()
          end
        end
      else:
        thread_flag_1903 = 2
      end
      if (thread_flag_1903 == 2):
        $ 1931 "Else" "noBreak"
        $ 1932 "exeption"
        $ 1933 "error"
        $ 1935 "OBJ_Brc_OK≔ False "
        global OBJ_Brc_OK=  False
      end
      $ 1936 "Set GRP_3F_Decap=Off"
      set_standard_digital_out(3, False)
      $ 1937 "Set GRP_3F_Enable=Off"
      set_standard_digital_out(4, False)
      $ 1938 "Set OTriggerBarcode=Off"
      write_output_boolean_register(1, False)
    elif (15 == switch_1):
      $ 1939 "Case 15"
      $ 1940 "Detect"
      $ 1941 "Action_Info≔'detect'"
      global Action_Info="detect"
    elif (30 == switch_1):
      $ 1942 "Case 30"
      $ 1943 "Shake"
      $ 1944 "Action_Info≔'shake'"
      global Action_Info="shake"
      $ 1945 "do_transition(pose_trans(FRM_Reference, PSE_T), keep_rxry=OBJ_Picked)"
      do_transition( pose_trans (FRM_Reference, PSE_T), keep_rxry=OBJ_Picked)
      $ 1946 "If PSE_A_H≠PSE_Z"
      if (PSE_A_H != PSE_Z):
        $ 1947 "If JNT_Q≠JNT_Z"
        if (JNT_Q != JNT_Z):
          $ 1948 "movej(get_inverse_kin(pose_trans(FRM_Reference, PSE_A_H), qnear=JNT_Q), r=0.050)"
          movej(get_inverse_kin( pose_trans (FRM_Reference, PSE_A_H), qnear=JNT_Q), r=0.050)
        else:
          $ 1949 "Else" "noBreak"
          $ 1950 "movej(pose_trans(FRM_Reference, PSE_A_H), r=0.050)"
          movej( pose_trans (FRM_Reference, PSE_A_H), r=0.050)
        end
      end
      $ 1951 "If PSE_A≠PSE_Z"
      if (PSE_A != PSE_Z):
        $ 1952 "If JNT_Q≠JNT_Z"
        if (JNT_Q != JNT_Z):
          $ 1953 "movej(get_inverse_kin(pose_trans(FRM_Reference, PSE_A), qnear=JNT_Q), r=0.020)"
          movej(get_inverse_kin( pose_trans (FRM_Reference, PSE_A), qnear=JNT_Q), r=0.020)
        else:
          $ 1954 "Else" "noBreak"
          $ 1955 "movej(pose_trans(FRM_Reference, PSE_A), r=0.020)"
          movej( pose_trans (FRM_Reference, PSE_A), r=0.020)
        end
      end
      $ 1956 "MoveL"
      $ 1957 "If PSE_T_H≠PSE_Z"
      if (PSE_T_H != PSE_Z):
        $ 1958 "PSE_T_H" "breakAfter"
        movel(pose_trans(FRM_Reference, PSE_T_H), a=0.5, v=0.4, r=0.01)
      end
      $ 1959 "PSE_T" "breakAfter"
      movel(pose_trans(FRM_Reference, PSE_T), a=0.08, v=0.12)
      $ 1960 "EXTT"
      $ 1961 "Comment"
      # Comment
      $ 1962 "MoveJ"
      $ 1963 "Waypoint_54" "breakAfter"
      movej(get_inverse_kin(Waypoint_54_p, qnear=Waypoint_54_q), a=1.3962634015954636, v=1.0471975511965976)
      $ 1964 "MoveJ"
      $ 1965 "Waypoint_77" "breakAfter"
      movej(get_inverse_kin(Waypoint_77_p, qnear=Waypoint_77_q), a=1.3962634015954636, v=1.0471975511965976)
      $ 1966 "MoveJ"
      $ 1967 "Waypoint_83" "breakAfter"
      movej(get_inverse_kin(Waypoint_83_p, qnear=Waypoint_83_q), a=1.3962634015954636, v=1.0471975511965976)
      $ 1968 "MoveJ"
      $ 1969 "Waypoint_84" "breakAfter"
      movej(get_inverse_kin(Waypoint_84_p, qnear=Waypoint_84_q), a=1.3962634015954636, v=1.0471975511965976)
      $ 1970 "If PSE_R_H≠PSE_Z"
      if (PSE_R_H != PSE_Z):
        $ 1971 "PSE_R" "breakAfter"
        movel(pose_trans(FRM_Reference, PSE_R), a=0.5, v=0.4, r=0.01)
        $ 1972 "PSE_R_H" "breakAfter"
        movel(pose_trans(FRM_Reference, PSE_R_H), a=0.5, v=0.4)
      else:
        $ 1973 "Else" "noBreak"
        $ 1974 "PSE_R" "breakAfter"
        movel(pose_trans(FRM_Reference, PSE_R), a=0.5, v=0.4)
      end
    elif (31 == switch_1):
      $ 1975 "Case 31"
      $ 1976 "Action_Info≔'Pick_Vial'"
      global Action_Info="Pick_Vial"
      $ 1977 "Pick_Vial"
      # begin: URCap Program Node
      #   Source: Robotiq_Grippers, 3.17.0.105337, Robotiq Inc.
      #   Type: Gripper
      $ 1978 "Gripper Open (1)"
      if not(gripper_connected[0]):
        popup("Gripper 1 must be connected to run this program.", "No connection", False, True, True)
      end
      if not(rq_is_gripper_activated("1")):
        popup("Gripper 1 is not activated. Go to Installation tab > Gripper to activate it and run the program again.", "Not activated", False, True, True)
      end
      rq_set_pos_spd_for(0, 82, 71, "1")
      rq_wait_pos_spe_for_request(0, 82, 71, "1")
      rq_go_to("1")
      rq_wait("1")
      # end: URCap Program Node
      $ 1979 "MoveJ"
      $ 1980 "Vial_above_1" "breakAfter"
      movej(get_inverse_kin(Vial_above_1_p, qnear=Vial_above_1_q), a=0.5235987755982988, v=0.4363323129985824, r=0.05)
      $ 1981 "MoveL"
      $ 1982 "Vial_pick_poi_1" "breakAfter"
      movel(Vial_pick_poi_1_p, a=0.5, v=0.1)
      # begin: URCap Program Node
      #   Source: Robotiq_Grippers, 3.17.0.105337, Robotiq Inc.
      #   Type: Gripper
      $ 1983 "Gripper Close (1)"
      if not(gripper_connected[0]):
        popup("Gripper 1 must be connected to run this program.", "No connection", False, True, True)
      end
      if not(rq_is_gripper_activated("1")):
        popup("Gripper 1 is not activated. Go to Installation tab > Gripper to activate it and run the program again.", "Not activated", False, True, True)
      end
      rq_set_pos_spd_for(255, 71, 84, "1")
      rq_wait_pos_spe_for_request(255, 71, 84, "1")
      rq_go_to("1")
      rq_wait("1")
      # end: URCap Program Node
      $ 1984 "MoveL"
      $ 1985 "Waypoint_86" "breakAfter"
      movel(Waypoint_86_p, a=0.5, v=0.1, r=0.05)
      $ 1986 "Home (Safe)"
      movej([-1.2302089344500047, -1.2969853503591224, -1.875639182904262, -1.539621866126728, 1.5731943360401213, -2.80099559440227], a=1.3962634015954636, v=1.0471975511965976)
    elif (32 == switch_1):
      $ 1987 "Case 32"
      $ 1989 "decap_Vial"
      $ 1990 "Set GRP_3F_Open=On"
      set_standard_digital_out(5, True)
      $ 1991 "MoveJ"
      $ 1992 "Waypoint_87" "breakAfter"
      movej(get_inverse_kin(Waypoint_87_p, qnear=Waypoint_87_q), a=0.5235987755982988, v=0.4363323129985824)
      $ 1993 "MoveL"
      $ 1994 "Vial_3FG_plac_1" "breakAfter"
